(* IEC 61131-3 sources: daoli-st-library/DL_Process (part 26) *)

(* ---- FB_DL_ChamberPumpDownProfile.st ---- *)
//==============================================================================
// 功能块：FB_DL_ChamberPumpDownProfile ｜ 中文名称：腔体抽气曲线包络监视
// 所属子库：DL_Process ｜ 版本：v1.0.0 ｜ 兼容：CODESYS V3.5+ / TwinCAT 3 / 汇川 InoProShop
// 功能描述：真空腔体抽气过程包络监视——启动时锁定基线压力，以指数衰减
//           包络为参照：包络上界 p_env(t) = fBasePa x EXP(-t/tau 包络)，
//           实测压力高于上界（衰减慢于包络）持续 tSlopeTimeout → 抽速
//           异常早停（bPumpAbortReq 锁存）；滚动窗内压力样本统计（窗口
//           极差）用于判「压力停滞」（极差 < 停滞阈且未达目标真空，同
//           样归入抽速异常）。达目标真空 → 抽气完成放行（信息级）。
//           斜率判据与窗统计互为冗余：一条失效另一条仍可兜住（如压力
//           缓慢泄漏时斜率判据先报，压力卡死时停滞判据先报）。
// 遗留假设（R95 代理阈值三句）：① 代理值 = fCycleTimeS 组态扫描周期
//           [秒]（包络时间基量）；② 覆盖 0.001~0.1 秒任务周期范围；
//           ③ 覆盖不到的区间由调用方按实际任务周期重设该引脚负责，
//           该假设挂编译验证债。
// 开源溯源 (Origin)：道莅原创实现（参考真空系统抽气曲线与抽速异常判定工程惯例 分类与参数域）
// 单位表：压力[帕] / 目标真空[帕] / 包络时间常数[秒] / 时间[ms] /
//         停滞阈[帕] / 极差[帕] / 扫描周期[秒] / 样本计数[次]
// 错误码表：16#0005_01F2 信息级（抽气完成：达目标真空放行，不置
//           bError）/ 16#0005_01F3 信息级（包络逼近预警：实测压力进入
//           包络上界 1.2 倍预警带，不置 bError）/ 16#0005_0330 故障级
//           （组态非法：目标/包络/阈值域、时间窗 <= 0 或任一输入非
//           有限，置 bError）/ 16#0005_0331 故障级（抽速异常早停：斜率
//           判据或停滞判据确认，bPumpAbortReq 锁存，置 bError——该场景
//           不可由 0330 的组态类判据观测，属工艺过程独立域）/
//           16#0005_0332 故障级兜底（状态机落 ELSE，置 bError）
// 状态机：E_DL_PumpDownState（五态：eIdle=0 / ePumping=10 / eDone=20 /
//           eAbort=30 / eFault=99），CASE 含 ELSE 兜底，ELSE 置 0332 并
//           撤早停请求外的全部输出
// 边界行为：① 组态非法 → 故障态锁存，bReset 复位；② 启动拍锁定基线
//           （基线取当拍实测，非魔法数）；③ 压力非有限 → 归入抽速异常
//           域早停（0331 复用，R90：传感器数据不可信时早停为安全侧）；
//           ④ 早停锁存至 bReset；⑤ 未启动/故障态早停请求撤零并
//           bValid := FALSE（空闲态不挂请求，防误触发停泵）；⑥ 窗口
//           样本环形缓存 8 点，满窗前停滞判据不生效（样本不足不判）。
// 修订历史：v1.0.0 2026-11-17 首版（R24 派单 · ROADMAP P1 §708）
//==============================================================================

(*------------------------------------------------------------------------------
 * 枚举: E_DL_PumpDownState（归属本功能块，同文件发布，全库唯一定义）
 * 含义: 抽气监视相位，每个成员在 CASE 中有且仅有一个标签。
 *-----------------------------------------------------------------------------*)
TYPE E_DL_PumpDownState :
(
    eIdle    := 0,   // 空闲：等启动沿 / Idle, awaiting start edge
    ePumping := 10,  // 抽气：包络与停滞双判据监视 / Pumping, envelope and stagnation dual monitoring
    eDone    := 20,  // 完成：达目标真空放行 / Done, target vacuum reached
    eAbort   := 30,  // 早停：抽速异常锁存 / Abort, pumping anomaly latched
    eFault   := 99   // 故障：组态非法/非法状态 / Fault, config or illegal state
);
END_TYPE

FUNCTION_BLOCK FB_DL_ChamberPumpDownProfile
VAR_INPUT
    bStart       : BOOL;                    // 启动请求 [—]，上升沿生效 / Start request, rising edge
    bReset       : BOOL;                    // 故障复位 [—]，上升沿清锁存 / Fault reset, rising edge clears latches
    fPressPa     : LREAL;                   // 腔压实测 [帕]（绝对压力） / Chamber pressure [Pa], absolute
    fTargetPa    : LREAL := 10.0;           // 目标真空 [帕]，须 > 0 / Target vacuum [Pa], must be > 0
    fTauEnvS     : LREAL := 60.0;           // 包络时间常数 [秒]，须 > 0 / Envelope time constant [s]
    fStagThreshPa: LREAL := 0.5;            // 停滞阈 [帕]（窗极差低于此判停滞） / Stagnation threshold [Pa]
    fSlopeMargin : LREAL := 1.2;            // 包络预警带倍数 [倍]（须 >= 1） / Envelope warning margin [ratio]
    tSlopeTimeout: TIME  := T#30S;          // 抽速异常确认窗 [ms]，须 > 0 / Anomaly confirm window [ms]
    fCycleTimeS  : LREAL := 0.01;           // 任务扫描周期 [秒]，须 > 0（R95 代理阈值） / Task scan cycle [s], must be > 0, R95 proxy
END_VAR
VAR_OUTPUT
    bPumpAbortReq : BOOL;                   // 抽速异常早停请求 [—]（锁存保持） / Pump-abort request, latched
    bPumpDownDone : BOOL;                   // 抽气完成 [—]（完成态电平） / Pump-down done, completion level
    fEnvPressPa   : LREAL;                  // 包络上界 [帕]（诊断出口） / Envelope ceiling [Pa], diagnostics outlet
    eState        : E_DL_PumpDownState;     // 相位出口 [—] / Phase outlet
    eErr          : UDINT;                  // 错误码，0 = 无错，码位 16#0005_01F2 起信息级、16#0005_0330 起故障级（分带见错误码表） / Error code, 0 = no error, band info/fault per the code table
    bError        : BOOL;                   // 故障级标志，仅故障级错误置位 / Fault-class flag, set only on fault-level codes
    bValid        : BOOL;                   // 输出可用标志 / Outputs usable flag
END_VAR
VAR
    fbSlope  : TON;                         // 抽速异常确认计时（每拍无条件刷新）[ms] / Anomaly confirm timer, refreshed unconditionally
    _eState  : E_DL_PumpDownState := E_DL_PumpDownState.eIdle; // 当前相位 / Current phase
    _bCfgBad : BOOL;                        // 组态非法锁存 / Illegal config latch
    _bAbortL : BOOL;                        // 早停锁存 / Abort latch
    _bInfoDone: BOOL;                       // 完成信息当拍标志 / Done info flag of this scan
    _bInfoWarn: BOOL;                       // 预警信息当拍标志 / Warning info flag of this scan
    _fBasePa : LREAL;                       // 启动基线压力 [帕] / Startup baseline pressure [Pa]
    _fElapsedS: LREAL;                      // 抽气累计时间 [秒] / Elapsed pumping time [s]
    _afWin   : ARRAY[0..7] OF LREAL;        // 滚动窗样本环形缓存 [帕] / Rolling-window sample ring [Pa]
    _nWinIdx : INT;                         // 环形缓存写指针 [次] / Ring write index [count]
    _nWinFill: INT;                         // 环形缓存已填数 [次] / Ring fill count [count]
    _bSlopeBad: BOOL;                       // 斜率判据电平（确认窗条件） / Slope-criterion level
    _bStagBad : BOOL;                       // 停滞判据电平（确认窗条件） / Stagnation-criterion level
    _bIllegal : BOOL;                       // 非法状态标志 / Illegal state flag
    _bInit    : BOOL := FALSE;              // 首扫标志，初值 FALSE 取非判定 / First-scan flag, tested negated
END_VAR
VAR CONSTANT
    DL_CPD_INF    : LREAL := 1.7976931348623157E308; // LREAL 幅值上限 / LREAL magnitude ceiling
    DL_CPD_EPS    : LREAL := 1.0E-6;        // 浮点判零容差 [帕] / Float zero tolerance [Pa]
    DL_CPD_WIN    : INT    := 8;            // 滚动窗容量 [次] / Rolling-window capacity [count]
    DL_CPD_ZERO   : LREAL := 0.0;           // 零值常量，避免裸字面量 [混合] / Zero constant, avoids a bare literal
END_VAR
VAR
    nI       : INT;                         // 极差统计循环索引 [次] / Range-statistics loop index
    fWinHi   : LREAL;                       // 窗内最大值 [帕] / Window maximum [Pa]
    fWinLo   : LREAL;                       // 窗内最小值 [帕] / Window minimum [Pa]
END_VAR

(*------------------------------------------------------------------------------
 * 段 1｜每拍预置：早停请求先撤（安全侧；锁存态在段 6 重置），标志预清零
 *      Abort request cleared first, flags pre-cleared
 *-----------------------------------------------------------------------------*)
bPumpAbortReq := FALSE;                  // 早停请求先撤（锁存态在段 6 重置） / Abort request cleared first
bPumpDownDone := FALSE;                  // 完成电平先清 / Done level cleared first
fEnvPressPa   := DL_CPD_ZERO;            // 包络出口每拍重算 / Envelope outlet recomputed
eErr   := 16#0000_0000;                  // 错误码每拍重算 / Error code recomputed
bError := FALSE;                         // 故障标志每拍重算 / Fault flag recomputed
bValid := FALSE;                         // 可用标志每拍重算 / Usable flag recomputed
_bInfoDone := FALSE;                     // 完成信息预清零 / Done info pre-cleared
_bInfoWarn := FALSE;                     // 预警信息预清零 / Warn info pre-cleared
_bIllegal  := FALSE;                     // 非法状态预清零 / Illegal flag pre-cleared

(*------------------------------------------------------------------------------
 * 段 2｜首扫初始化
 *      First-scan initialisation
 *-----------------------------------------------------------------------------*)
IF NOT _bInit THEN
    _eState  := E_DL_PumpDownState.eIdle; // 相位空闲起步 / Phase starts idle
    _bCfgBad := FALSE;                   // 组态锁存清零 / Config latch cleared
    _bAbortL := FALSE;                   // 早停锁存清零 / Abort latch cleared
    _fElapsedS := DL_CPD_ZERO;           // 累计时间清零 / Elapsed time cleared
    _nWinIdx := 0;                       // 写指针归零 / Write index reset
    _nWinFill := 0;                      // 已填数归零 / Fill count reset
    _bInit   := TRUE;                    // 首扫只做一次 / The first scan runs once
END_IF

(*------------------------------------------------------------------------------
 * 段 3｜组态防御闸：非有限（R79）+ 目标/包络/阈值/时间窗域
 *      Configuration defense gates
 *-----------------------------------------------------------------------------*)
IF (fTargetPa <> fTargetPa) OR (ABS(fTargetPa) > DL_CPD_INF)
   OR (fTauEnvS <> fTauEnvS) OR (ABS(fTauEnvS) > DL_CPD_INF)
   OR (fStagThreshPa <> fStagThreshPa) OR (ABS(fStagThreshPa) > DL_CPD_INF)
   OR (fSlopeMargin <> fSlopeMargin) OR (ABS(fSlopeMargin) > DL_CPD_INF)
   OR (fCycleTimeS <> fCycleTimeS) OR (ABS(fCycleTimeS) > DL_CPD_INF) THEN
    _bCfgBad := TRUE;                    // 非有限归组态非法锁存 / Non-finite folded into the config latch
END_IF
IF (NOT _bCfgBad) AND ((fTargetPa <= DL_CPD_EPS) OR (fTauEnvS <= DL_CPD_EPS)
   OR (fStagThreshPa <= DL_CPD_EPS) OR (fSlopeMargin < 1.0)
   OR (tSlopeTimeout <= T#0MS) OR (fCycleTimeS <= DL_CPD_EPS)) THEN
    _bCfgBad := TRUE;                    // 目标/包络/阈值/时间窗域非法锁存 / Target, envelope, threshold and window domains latched
END_IF
IF bReset THEN
    _bCfgBad := FALSE;                   // 复位清组态锁存 / Reset clears the config latch
    _bAbortL := FALSE;                   // 复位清早停锁存 / Reset clears the abort latch
END_IF

(*------------------------------------------------------------------------------
 * 段 4｜确认窗无条件刷新（R40：CASE 之外每拍必调）
 *      Confirm timer refreshed unconditionally per R40
 *-----------------------------------------------------------------------------*)
fbSlope(IN := (_eState = E_DL_PumpDownState.ePumping)
             AND (_bSlopeBad OR _bStagBad), PT := tSlopeTimeout); // 抽速异常确认窗 / Anomaly confirm window

(*------------------------------------------------------------------------------
 * 段 5｜相位机与双判据链（CASE 含 ELSE 兜底；状态改写只出现在分支判据内，R39）
 *      Phase machine and the dual-criteria chain
 *-----------------------------------------------------------------------------*)
CASE _eState OF

    E_DL_PumpDownState.eIdle:              // 空闲：启动沿且组态合法进抽气
        IF bStart AND (NOT _bCfgBad) THEN
            _fBasePa := fPressPa;          // 基线锁定（启动拍实测，非魔法数） / Baseline locked at start
            _fElapsedS := DL_CPD_ZERO;     // 累计时间归零 / Elapsed time reset
            _nWinIdx := 0;                 // 写指针归零 / Write index reset
            _nWinFill := 0;                // 已填数归零（满窗前停滞判据不生效） / Fill reset, stagnation inert before the full window
            _eState := E_DL_PumpDownState.ePumping; // 进抽气 / To pumping
        ELSIF bStart AND _bCfgBad THEN
            _eState := E_DL_PumpDownState.eFault; // 组态非法进故障 / Illegal config to fault
        END_IF

    E_DL_PumpDownState.ePumping:           // 抽气：包络/停滞双判据 + 目标判定
        IF _bCfgBad THEN
            _eState := E_DL_PumpDownState.eFault; // 组态漂移转故障 / Config drift, fault
        ELSIF fPressPa <= fTargetPa THEN
            _bInfoDone := TRUE;            // 达目标真空（信息级，拍 N 进入） / Target vacuum reached, info
            _eState := E_DL_PumpDownState.eDone; // 本拍转出：进完成 / To done
        ELSE
            _fElapsedS := _fElapsedS + fCycleTimeS; // 累计时间推进 [秒] / Elapsed time advanced
            IF (fPressPa <> fPressPa) OR (ABS(fPressPa) > DL_CPD_INF) THEN
                _bSlopeBad := TRUE;        // 腔压非有限归抽速异常域（传感器数据不可信，早停安全侧，0331 复用 R90） / Non-finite pressure folded into the anomaly domain
            ELSE
                fEnvPressPa := _fBasePa * EXP(-_fElapsedS / fTauEnvS); // 包络上界 [帕]，分母已闸 / Envelope ceiling, denominator gated
                _bSlopeBad := fPressPa > (fSlopeMargin * fEnvPressPa); // 斜率判据：衰减慢于包络 / Slope criterion: slower than the envelope
            END_IF
            _afWin[_nWinIdx] := fPressPa;  // 样本入环 / Sample into the ring
            _nWinIdx := (_nWinIdx + 1) MOD DL_CPD_WIN; // 写指针环形推进（模 8，归一安全） / Ring index advance, modulo-normalised
            IF _nWinFill < DL_CPD_WIN THEN
                _nWinFill := _nWinFill + 1; // 已填数推进 / Fill count advanced
            END_IF
            IF _nWinFill >= DL_CPD_WIN THEN
                fWinHi := _afWin[0];       // 窗极差统计起步 / Range statistics start
                fWinLo := _afWin[0];       // 窗极差统计起步 / Range statistics start
                FOR nI := 1 TO (DL_CPD_WIN - 1) DO
                    IF _afWin[nI] > fWinHi THEN
                        fWinHi := _afWin[nI]; // 窗内最大值 / Window maximum
                    END_IF
                    IF _afWin[nI] < fWinLo THEN
                        fWinLo := _afWin[nI]; // 窗内最小值 / Window minimum
                    END_IF
                END_FOR
                _bStagBad := (fWinHi - fWinLo) < fStagThreshPa; // 停滞判据：窗极差低于阈 / Stagnation: range below the threshold
            ELSE
                _bStagBad := FALSE;        // 样本不足不判停滞（边界行为⑥） / Sample insufficient, no stagnation verdict
            END_IF
            IF fbSlope.Q THEN
                _bAbortL := TRUE;          // 抽速异常确认，早停锁存（拍 N 进入） / Anomaly confirmed, abort latched
                _eState := E_DL_PumpDownState.eAbort; // 本拍转出：进早停 / To abort
            END_IF
        END_IF

    E_DL_PumpDownState.eDone:              // 完成：等启动撤销回空闲（同拍重启防抖）
        IF NOT bStart THEN
            _eState := E_DL_PumpDownState.eIdle; // 回空闲 / Back to idle
        END_IF

    E_DL_PumpDownState.eAbort:             // 早停：请求锁存保持，bReset 才解除
        IF bReset AND (NOT _bCfgBad) THEN
            _bAbortL := FALSE;             // 复位清早停锁存 / Reset clears the abort latch
            _eState := E_DL_PumpDownState.eIdle; // 回空闲 / Back to idle
        END_IF

    E_DL_PumpDownState.eFault:             // 故障：复位沿且组态恢复回空闲
        IF bReset AND (NOT _bCfgBad) THEN
            _eState := E_DL_PumpDownState.eIdle; // 回空闲 / Back to idle
        END_IF

    ELSE                                   // 非法状态兜底（R21：CASE 必带 ELSE）
        _bIllegal := TRUE;                 // 标记非法状态 / Flag the illegal state
        _eState := E_DL_PumpDownState.eFault; // 回故障态 / Back to fault
END_CASE

IF (_eState = E_DL_PumpDownState.ePumping) AND (_fElapsedS > DL_CPD_EPS)
   AND (fPressPa > (fSlopeMargin * fEnvPressPa)) THEN
    _bInfoWarn := TRUE;                    // 包络逼近预警带（信息级） / Envelope approach warning, info
END_IF

(*------------------------------------------------------------------------------
 * 段 6｜码位出口与放行（故障级码 3 行内置 bError，R45/R101 配对）
 *      Code outlet and release, fault codes paired with bError
 *-----------------------------------------------------------------------------*)
IF _bIllegal THEN
    eErr   := 16#0005_0332;                // 故障级：状态机兜底 / Fault: state machine fallback
    bError := TRUE;                        // 置故障标志 / Raise the fault flag
ELSIF _bCfgBad THEN
    eErr   := 16#0005_0330;                // 故障级：组态非法 / Fault: illegal configuration
    bError := TRUE;                        // 置故障标志 / Raise the fault flag
ELSIF _bAbortL THEN
    eErr   := 16#0005_0331;                // 故障级：抽速异常早停锁存 / Fault: pumping anomaly, abort latched
    bError := TRUE;                        // 置故障标志 / Raise the fault flag
ELSIF _bInfoWarn THEN
    eErr := 16#0005_01F3;                  // 信息级：包络逼近预警 / Info: envelope approach warning
ELSIF _bInfoDone THEN
    eErr := 16#0005_01F2;                  // 信息级：抽气完成放行 / Info: pump-down done
END_IF

bPumpAbortReq := _bAbortL;               // 早停请求出口 = 锁存量（R99，空闲态不挂请求） / Abort outlet equals the latch
bPumpDownDone := (_eState = E_DL_PumpDownState.eDone); // 完成电平挂状态量 / Done level bound to the state
bValid := (NOT bError) AND (_eState <> E_DL_PumpDownState.eIdle); // 空闲/故障输出不可用 / Outputs unusable in idle or fault
eState := _eState;                       // 相位出口 / Phase outlet
END_FUNCTION_BLOCK

(* ---- FB_DL_ChamberPurgeDry.st ---- *)
(*
  FB_DL_ChamberPurgeDry  —  腔体干燥吹扫顺控 / Chamber purge and dry sequence control
  分类 Category : DL_Process
  码位 Code     : 16#06_0_82
  版本 Version  : 1.0.1
  溯源 Source   : OSCAT Building 语义借鉴 · clean-room 实现，仅借分类/参数域/命名，未复制源码
  修改记录 Hist : v1.0.1 2026-11-23 R75 修复——FC_DL_DewPointCalc 调用补
                  uErrorId / fVaporPa / bInRange 三出参显式回执（R73 零回执
                  挂账点修，与 VaporPressureSat 族回执口径对齐），bInRange
                  并入有效判据，主顺控逻辑零改动
  功能 Function : 1) 露点判据收敛：吹扫 → 静置 → 复测 三态循环，直到复测露点低于目标；
                  2) 三段计时各用独立 TON，且每段 IN := (在相) AND NOT ton.Q 自复位（FB33-2 硬判据）；
                  3) 复测未收敛不无限等待，超过 nMaxRetry 次即转超时态并报码。
  边界 Boundary : ① 露点入参先过有限性与物理域闸（RH 0~100 %、温度 −40~120 °C），域外不出结论；
                  ② 吹扫/静置/复测计时用三实例分段 TON，每段自复位；
                  ③ 复测超次即超时升级，不得延续吹扫无限等待；
                  ④ 超时/故障三行同向：吹扫阀关 → 干燥气阀关 → 进度标志 FALSE。
  依赖 Depends  : FC_DL_DewPointCalc（露点换算，每拍无条件调用）

  码表 Error codes（本件子码步进 16#10，避让邻件码位）:
    16#0002_0682 故障级：露点入参域外或露点函数返回无效（域闸锁存，输入恢复后自解）
    16#0002_0692 故障级：计时参数为 0 或重试上限 < 1（组态闸锁存，需 bReset 清除）
    16#0002_06A2 信息级：复测超次转超时（不置 bError，仅提示）
*)

TYPE E_DL_PurgeDryPhase :
(
    eIdle      := 0,   // 空闲 / Idle
    ePurge     := 10,  // 吹扫段 / Purge stage
    eSoak      := 20,  // 静置段 / Soak stage
    eRemeasure := 30,  // 复测段 / Re-measure stage
    eDone      := 40,  // 干燥达标 / Dry target reached
    eTimeout   := 50,  // 复测超次超时 / Retry timeout
    eFault     := 90   // 故障锁定 / Fault locked
);
END_TYPE

FUNCTION_BLOCK FB_DL_ChamberPurgeDry
VAR_INPUT
    bEnable        : BOOL;                        // 总使能，FALSE 回空闲关阀 / Master enable
    bStart         : BOOL;                        // 启动，上升沿有效 / Start, rising edge
    bReset         : BOOL;                        // 复位，上升沿清故障与超时 / Reset, clears fault and timeout
    fTempC         : REAL;                        // 腔体干球温度 [degC]，域 −40~120 / Chamber dry-bulb temperature [degC]
    fRhPct         : REAL;                        // 腔体相对湿度 [%]，域 0~100 / Chamber relative humidity [%]
    fDewTargetC    : REAL := -20.0;               // 露点目标 [degC]，复测低于此值判达标 / Dew point target [degC]
    fDewHystC      : REAL := 2.0;                 // 露点达标迟滞 [degC]，防边界抖动 / Dew point hysteresis [degC]
    tPurgeTime     : TIME := T#60S;               // 吹扫段时长 [ms]，域 > 0 / Purge stage duration
    tSoakTime      : TIME := T#30S;               // 静置段时长 [ms]，域 > 0 / Soak stage duration
    tRemeasureTime : TIME := T#20S;               // 复测段时长 [ms]，域 > 0 / Re-measure stage duration
    tDewSampleTime : TIME := T#500MS;             // 露点采样节拍 [ms]，自复位心跳 / Dew sample tick, self-resetting
    nMaxRetry      : INT := 5;                    // 最大复测次数 [次]，域 >= 1 / Max re-measure count
END_VAR
VAR_OUTPUT
    bPurgeValve    : BOOL;                        // 吹扫进气阀 [开关] / Purge inlet valve
    bDryAirValve   : BOOL;                        // 干燥气补充阀 [开关] / Dry air makeup valve
    bExhaustValve  : BOOL;                        // 排气阀 [开关] / Exhaust valve
    fDewNowC       : REAL;                        // 当前露点 [degC]，采样节拍刷新 / Current dew point [degC]
    bDewValid      : BOOL;                        // 露点有效标志 / Dew point valid flag
    nRetry         : INT;                         // 已复测次数 [次] / Re-measure count
    bInProgress    : BOOL;                        // 顺控进行中 / Sequence in progress
    bDone          : BOOL;                        // 达标完成（保持型）/ Dry done, level held
    bTimeout       : BOOL;                        // 超时标志（保持型）/ Timeout flag, level held
    bError         : BOOL;                        // 故障标志，与故障级码配对 / Fault flag paired with fault codes
    uErrorId       : UDINT;                       // 事件码，0 = 无事件 / Event code, 0 = none
    eStateOut      : E_DL_PurgeDryPhase;          // 状态机当前态，段尾单点映射 / Phase mapped at tail
END_VAR
VAR
    _eState        : E_DL_PurgeDryPhase := E_DL_PurgeDryPhase.eIdle;  // 内部状态 / Internal state
    rtrStart       : R_TRIG;                      // 启动沿 / Start edge
    rtrReset       : R_TRIG;                      // 复位沿 / Reset edge
    tonPurge       : TON;                         // 吹扫段计时（自复位）/ Purge stage timer, self-resetting
    tonSoak        : TON;                         // 静置段计时（自复位）/ Soak stage timer, self-resetting
    tonRemeasure   : TON;                         // 复测段计时（自复位）/ Re-measure stage timer
    tonDewTick     : TON;                         // 露点采样心跳（自复位）/ Dew sample tick, self-resetting
    fDewCalcC      : REAL;                        // 露点函数返回暂存 [degC] / Dew point function result
    fDewHoldC      : REAL;                        // 采样节拍锁存露点 [degC] / Latched dew point at tick
    bInputOk       : BOOL;                        // 露点入参域闸结果 / Dew input domain result
    bCfgOk         : BOOL;                        // 计时/重试组态合法 / Timer and retry configuration valid
    bConverged     : BOOL;                        // 复测收敛标志 / Convergence flag
    uFault         : UDINT;                       // 锁存故障码 / Latched fault code
    uInfo          : UDINT;                       // 信息级码 / Information code
    uDewErr        : UDINT;                       // 露点函数回执码（v1.0.1 新增接收）/ Dew point FC receipt, new in v1.0.1
    fVaporPaBuf    : REAL;                        // 露点函数水汽压回执 [Pa]（v1.0.1 新增接收，诊断）/ Dew point FC vapor pressure receipt [Pa]
    bDewInRange    : BOOL;                        // 露点函数域内回执 [-]（v1.0.1 新增接收）/ Dew point FC in-range receipt
END_VAR
VAR CONSTANT
    DL_PD_TMIN     : REAL := -40.0;               // 温度有效域下限 [degC] / Temperature domain low [degC]
    DL_PD_TMAX     : REAL := 120.0;               // 温度有效域上限 [degC] / Temperature domain high [degC]
    DL_PD_RHMIN    : REAL := 0.0;                 // 湿度有效域下限 [%] / Humidity domain low [%]
    DL_PD_RHMAX    : REAL := 100.0;               // 湿度有效域上限 [%] / Humidity domain high [%]
END_VAR

(* === 段 0 · 实例刷新（无条件周期调用，自复位节拍）=== *)
rtrStart(CLK := bStart);                          // 每拍刷新启动沿
rtrReset(CLK := bReset);                          // 每拍刷新复位沿
tonPurge(IN := (_eState = E_DL_PurgeDryPhase.ePurge) AND (NOT tonPurge.Q), PT := tPurgeTime);      // 自复位
tonSoak(IN := (_eState = E_DL_PurgeDryPhase.eSoak) AND (NOT tonSoak.Q), PT := tSoakTime);           // 自复位
tonRemeasure(IN := (_eState = E_DL_PurgeDryPhase.eRemeasure) AND (NOT tonRemeasure.Q), PT := tRemeasureTime); // 自复位
tonDewTick(IN := NOT tonDewTick.Q, PT := tDewSampleTime);                                            // 采样心跳自复位

(* === 段 1 · 域闸：入参有限性 + 物理域，域外不出结论 === *)
bInputOk := (fTempC = fTempC) AND (fRhPct = fRhPct)                          // NaN 自反判据
            AND (ABS(fTempC) < 1.0E30) AND (ABS(fRhPct) < 1.0E30)            // Inf 上限兜底
            AND (fTempC >= DL_PD_TMIN) AND (fTempC <= DL_PD_TMAX)            // 温度物理域闸
            AND (fRhPct >= DL_PD_RHMIN) AND (fRhPct <= DL_PD_RHMAX);         // 湿度物理域闸
fDewCalcC := FC_DL_DewPointCalc(fTempC := fTempC, fRhPct := fRhPct,
                                uErrorId => uDewErr, fVaporPa => fVaporPaBuf,
                                bInRange => bDewInRange);                   // 露点换算每拍无条件调用 + 三出参回执（v1.0.1）
IF bInputOk AND bDewInRange AND (fDewCalcC = fDewCalcC) AND (ABS(fDewCalcC) < 1.0E30) THEN   // 域内回执并入判据（v1.0.1）
    IF tonDewTick.Q THEN
        fDewHoldC := fDewCalcC;                   // 采样节拍到时锁存露点（每 N 时间采一次）
        bDewValid := TRUE;                        // 露点有效
    END_IF
ELSE
    bDewValid := FALSE;                           // 域外：露点无效，不清零旧值（保持诊断可读）
END_IF
bCfgOk := (tPurgeTime > T#0MS) AND (tSoakTime > T#0MS) AND (tRemeasureTime > T#0MS)
          AND (tDewSampleTime > T#0MS) AND (nMaxRetry >= 1);                 // 计时与重试组态闸
IF NOT bCfgOk THEN
    uFault := 16#0002_0692;                       // 故障级：计时参数为 0 或重试上限非法
END_IF
IF NOT bInputOk THEN
    uFault := 16#0002_0682;                       // 故障级：露点入参域外（输入恢复后段 2 自解）
END_IF
IF bInputOk AND bCfgOk THEN
    IF uFault = 16#0002_0682 THEN
        uFault := 16#0000;                        // 输入恢复即自解域闸故障（复位路径可达）
    END_IF
END_IF
IF rtrReset.Q AND bCfgOk THEN
    uFault := 16#0000;                            // 复位沿清锁存（组态已合法才允许）
END_IF

(* === 段 2 · 主状态机（ENUM + CASE，含 ELSE 兜底）=== *)
CASE _eState OF
E_DL_PurgeDryPhase.eIdle :
    nRetry := 0;                                  // 新一轮复测计数清零
    bDone := FALSE;                               // 完成标志复位
    bTimeout := FALSE;                            // 超时标志复位
    bConverged := FALSE;                          // 收敛标志复位
    uInfo := 16#0000;                             // 信息码清零（条件不满足则保持 0）
    IF uFault = 16#0002_0692 THEN
        _eState := E_DL_PurgeDryPhase.eFault;     // 组态故障优先拦截
    ELSIF rtrStart.Q THEN
        _eState := E_DL_PurgeDryPhase.ePurge;     // 本拍进入吹扫相
    END_IF

E_DL_PurgeDryPhase.ePurge :
    IF tonPurge.Q THEN
        _eState := E_DL_PurgeDryPhase.eSoak;      // 本拍行为：吹扫到时长，拍末转静置
    END_IF

E_DL_PurgeDryPhase.eSoak :
    IF tonSoak.Q THEN
        _eState := E_DL_PurgeDryPhase.eRemeasure; // 静置到时长，转复测相
    END_IF

E_DL_PurgeDryPhase.eRemeasure :
    IF tonRemeasure.Q THEN
        bConverged := bDewValid AND (fDewHoldC <= (fDewTargetC - fDewHystC));   // 露点低于目标减迟滞才判收敛
        nRetry := nRetry + 1;                     // 复测次数累加
        IF bConverged THEN
            _eState := E_DL_PurgeDryPhase.eDone;  // 收敛：转达标态
            bDone := TRUE;                        // 置位型：完成标志，段尾不清零
        ELSIF nRetry >= nMaxRetry THEN
            _eState := E_DL_PurgeDryPhase.eTimeout;   // 超次：超时升级，不无限等待
            bTimeout := TRUE;                     // 置位型：超时标志
            uInfo := 16#0002_06A2;                // 信息级：复测超次（不置 bError）
        ELSE
            _eState := E_DL_PurgeDryPhase.ePurge; // 未收敛且余次：回吹扫再循环
        END_IF
    END_IF

E_DL_PurgeDryPhase.eDone :
    bDone := TRUE;                                // 达标保持直到复位或再启动
    IF rtrStart.Q OR rtrReset.Q THEN
        _eState := E_DL_PurgeDryPhase.eIdle;      // 再启动/复位回空闲
    END_IF

E_DL_PurgeDryPhase.eTimeout :
    bTimeout := TRUE;                             // 超时标志保持，等人为处理
    IF rtrReset.Q THEN
        bTimeout := FALSE;                        // 复位沿解除超时（可到达的解除路径）
        uInfo := 16#0000;                         // 信息码同步清除
        _eState := E_DL_PurgeDryPhase.eIdle;
    END_IF

E_DL_PurgeDryPhase.eFault :
    IF (uFault = 16#0000) THEN
        _eState := E_DL_PurgeDryPhase.eIdle;      // 故障已解锁回空闲
    END_IF

ELSE
    _eState := E_DL_PurgeDryPhase.eFault;         // 非法状态拦截
    uFault := 16#0002_0692;                       // 故障级：相 ID 越界（枚举兜底路径）
END_CASE
IF NOT bEnable THEN
    _eState := E_DL_PurgeDryPhase.eIdle;          // 失能最高优先回空闲
    bInProgress := FALSE;                         // 进度标志随之为 FALSE
END_IF

(* === 段 3 · 输出映射（安全三行同向：阀门关 → 露点值 → 进度判据）=== *)
bPurgeValve   := (_eState = E_DL_PurgeDryPhase.ePurge);      // 吹扫阀仅吹扫相开
bDryAirValve  := (_eState = E_DL_PurgeDryPhase.ePurge) OR (_eState = E_DL_PurgeDryPhase.eSoak);  // 干燥气随吹扫/静置
bExhaustValve := (_eState = E_DL_PurgeDryPhase.ePurge) OR (_eState = E_DL_PurgeDryPhase.eSoak)
                 OR (_eState = E_DL_PurgeDryPhase.eRemeasure);   // 排气阀复测相亦开
IF (_eState = E_DL_PurgeDryPhase.eTimeout) OR (_eState = E_DL_PurgeDryPhase.eFault)
   OR (_eState = E_DL_PurgeDryPhase.eIdle) THEN
    bPurgeValve := FALSE;                         // 超时/故障/空闲：吹扫阀强制关
    bDryAirValve := FALSE;                        // 干燥气阀强制关
    bExhaustValve := FALSE;                       // 排气阀强制关
END_IF
fDewNowC := fDewHoldC;                            // 露点输出取采样锁存值
bInProgress := (_eState = E_DL_PurgeDryPhase.ePurge) OR (_eState = E_DL_PurgeDryPhase.eSoak)
               OR (_eState = E_DL_PurgeDryPhase.eRemeasure);   // 进度判据与阀门同向
bError := (uFault <> 16#0000);                    // 故障标志仅由故障级码置位（R45 配对）
IF bError THEN
    uErrorId := uFault;                           // 故障级优先上报
ELSE
    uErrorId := uInfo;                            // 否则上报信息级码
END_IF
eStateOut := _eState;                             // 输出枚举段尾单点映射（N2 规则）
END_FUNCTION_BLOCK

(* ---- FB_DL_ChamberTempUnitBank.st ---- *)
(*
  ==================================================================
  组件名 Component  : FB_DL_ChamberTempUnitBank
  分类   Category   : DL_Process
  版本   Version    : 1.0.0
  功能   Purpose    : 多腔室温标统一换算行。批量把 1..8 个腔室的温度实测值从
                      源温标（摄氏 / 华氏 / 开尔文）换算到目标温标，出口逐通道
                      结果、逐通道有效性掩码与统计计数。内核为「先归一到摄氏、
                      再由摄氏展开到目标温标」两段式，六种换向共用同一对归一 /
                      展开函数体，不存在重复公式分支。
  溯源   Origin     : 温标换算为公开物理定义（0 摄氏度 = 273.15 开尔文 = 32 华氏度，
                      华氏步长为摄氏的 1.8 倍）；本件为 clean-room 实现，仅借鉴来源
                      分类与参数域组织（来源标签 roadmap-p2-chamber），道莅原创设计，
                      未复制任何闭源代码行。
  平台   Platform   : 纯 IEC 61131-3（REAL / WORD / SHL 常量移位，无私有库）
  作者   Author     : 道莅代码库 · PLC 编程专家（R55）
  ------------------------------------------------------------------
  边界 Boundary     :
                      一 本件只做单位换算与有效性标记，不判工艺超温、不做滤波、不做报警；
                      二 非有限输入不穿透出口：该通道保持上拍值并置无效位；
                      三 结果低于目标温标绝对零度时按 bClampAbsZero 钳到绝对零点并置无效位；
                      四 通道游标经回钳 1..8，掩码位移量 0..7 由数组边界与循环上界共同证明；
                      五 无全局变量、无外部变量声明、无物理地址寻址。
  输出契约 Output contract:
                      afTempOut 逐通道结果；序号大于 nChamberCount 的通道保持上拍值不清零；
                      wInvalidMask 位 i-1 对应通道 i，自证向量：仅通道 1 无效 → 16#0001，
                      仅通道 8 无效 → 16#0080；
                      故障级成因 eUnitBad 与 bError 配对（R45），信息级成因永不置 bError。
  修订记录 Revision  :
    2026-11-20  v1.0.0  R55 首版（批 1 · 序号 4）
  ==================================================================
*)

TYPE E_DL_TempUnit :
(
    eCelsius    := 0,   // 摄氏度 [摄氏度] / degree Celsius
    eFahrenheit := 10,  // 华氏度 [华氏度] / degree Fahrenheit
    eKelvin     := 20   // 开尔文 [开尔文] / Kelvin
);
END_TYPE

TYPE E_DL_TubCause :
(
    eNone       := 0,   // 无成因 / no cause
    eUnitBad    := 1,   // 温标枚举非法（故障级，与 bError 配对）/ illegal temperature unit enumeration, a fault paired with bError
    eCountBad   := 2,   // 通道数越域已回钳（信息级）/ channel count out of domain and clamped, informational
    eChanBad    := 3,   // 存在非有限通道，已保持上拍值（信息级）/ non-finite channels present and held at the last value, informational
    eAbsZero    := 4    // 结果低于绝对零度已钳位（信息级）/ result below absolute zero and clamped, informational
);
END_TYPE

FUNCTION_BLOCK FB_DL_ChamberTempUnitBank
VAR_INPUT
    bEnable        : BOOL := TRUE;           // 使能，失能时全部通道保持上拍值 [-] / enable, all channels hold their last value when disabled
    bReset         : BOOL := FALSE;          // 复位上升沿清故障锁存与掩码 [-] / reset rising edge clears the fault latch and the mask
    eUnitIn        : E_DL_TempUnit := E_DL_TempUnit.eCelsius;    // 源温标 [枚举] / source temperature unit [enum]
    eUnitOut       : E_DL_TempUnit := E_DL_TempUnit.eCelsius;    // 目标温标 [枚举] / target temperature unit [enum]
    nChamberCount  : INT := 8;               // 参与换算的腔室数 [个]，域 1..8 / participating channels [count], domain 1 to 8
    bClampAbsZero  : BOOL := TRUE;           // 真 = 低于绝对零度钳位，假 = 仅置无效位不改值 [-] / true clamps below absolute zero, false only flags
END_VAR
VAR_IN_OUT
    afTempIn       : ARRAY[1..8] OF REAL;    // 逐腔室温度输入 [源温标单位]，引用型入参由调用方持有 / per chamber temperature inputs in source unit, reference parameter owned by the caller
END_VAR
VAR_OUTPUT
    afTempOut      : ARRAY[1..8] OF REAL := [8(0.0)]; // 逐腔室换算结果 [目标温标单位] / per chamber converted results in target unit
    wInvalidMask   : WORD := 16#0000;        // 无效通道掩码，位 i-1 对应通道 i [-] / invalid channel mask, bit i minus one maps to channel i
    nValidCount    : INT := 0;               // 本拍有效通道数 [个] / valid channel count of this scan
    bAllValid      : BOOL := FALSE;          // 全部参与通道有效 [-] / all participating channels valid
    bAnyInvalid    : BOOL := FALSE;          // 存在无效通道 [-] / at least one invalid channel
    fSumOut        : REAL := 0.0;            // 有效通道结果之和 [目标温标单位] / sum of the valid converted results
    fAvgOut        : REAL := 0.0;            // 有效通道结果均值 [目标温标单位] / mean of the valid converted results
    eCause         : E_DL_TubCause := E_DL_TubCause.eNone; // 成因出口 [枚举] / cause outlet [enum]
    bError         : BOOL := FALSE;          // 故障锁存标志 [-] / fault latch flag
END_VAR
VAR
    rtReset        : R_TRIG;                 // 复位沿检测，段 0 无条件刷新 / reset edge detector, refreshed unconditionally in segment zero
    _eCause        : E_DL_TubCause := E_DL_TubCause.eNone;  // 内部成因，故障级锁存、信息级每拍重算 / internal cause, latched for faults and recomputed for information
    _bFault        : BOOL := FALSE;          // 故障锁存位（温标枚举非法）/ fault latch bit for an illegal unit enumeration
    _bInit         : BOOL := FALSE;          // 首扫初始化完成标志（R310）/ first scan initialisation flag
    _bUnitInOk     : BOOL := FALSE;          // 源温标枚举合法性 [-] / source unit enumeration validity
    _bUnitOutOk    : BOOL := FALSE;          // 目标温标枚举合法性 [-] / target unit enumeration validity
    _bChanOk       : BOOL := FALSE;          // 单通道输入有限性 [-] / single channel input finiteness
    _bResultOk     : BOOL := FALSE;          // 单通道结果有限性 [-] / single channel result finiteness
    _bChanBitBad   : BOOL := FALSE;          // 单通道无效位 [-] / single channel invalid bit
    _bAbsZeroHit   : BOOL := FALSE;          // 本拍出现绝对零度钳位 [-] / an absolute zero clamp occurred this scan
    _bChanNonFin   : BOOL := FALSE;          // 本拍出现非有限通道 [-] / a non-finite channel occurred this scan
    _bCountClamped : BOOL := FALSE;          // 通道数被回钳 [-] / the channel count was clamped
    _nUseCount     : INT := 0;               // 钳定后的参与通道数 [个] / clamped participating channel count
    _nIdx          : INT := 0;               // 通道游标（1 起，回钳 1..8）[通道号] / channel cursor, one-based, clamped one through eight
    _fCelsius      : REAL := 0.0;            // 归一到摄氏度的中间量 [摄氏度] / intermediate normalised to Celsius
    _fResult       : REAL := 0.0;            // 展开到目标温标的中间量 [目标温标单位] / intermediate expanded to the target unit
    _fLowLimit     : REAL := 0.0;            // 目标温标绝对零度 [目标温标单位] / absolute zero in the target unit
    _fSum          : REAL := 0.0;            // 有效结果累加 [目标温标单位] / running sum of valid results
    _wMask         : WORD := 16#0000;        // 掩码累加器，每拍清零重建 / mask accumulator, rebuilt every scan
    _wBitOne       : WORD := 16#0001;        // 单位位常量，供常量移位使用 [-] / single bit constant for the shift
END_VAR
VAR CONSTANT
    DL_TUB_MAX        : INT := 8;            // 通道容量，同时也是游标回钳上界 [个] / channel capacity and cursor clamp upper bound
    DL_TUB_K_OFFSET   : REAL := 273.15;      // 摄氏与开尔文零点偏移 [开尔文] / zero offset between Celsius and Kelvin
    DL_TUB_F_RATIO    : REAL := 1.8;         // 华氏与摄氏步长比 [无量纲] / scale ratio between Fahrenheit and Celsius
    DL_TUB_F_OFFSET   : REAL := 32.0;        // 华氏零点偏移 [华氏度] / zero offset of Fahrenheit
    DL_TUB_ABS_C      : REAL := -273.15;     // 摄氏绝对零度 [摄氏度] / absolute zero in Celsius
    DL_TUB_ABS_F      : REAL := -459.67;     // 华氏绝对零度 [华氏度] / absolute zero in Fahrenheit
    DL_TUB_ABS_K      : REAL := 0.0;         // 开尔文绝对零度 [开尔文] / absolute zero in Kelvin
    DL_TUB_ABS_MARGIN : REAL := 0.01;        // 绝对零度容差带，吸收换算舍入 [目标温标单位] / absolute zero tolerance absorbing rounding
    DL_TUB_MASK_NONE  : WORD := 16#0000;     // 空掩码常量 [-] / empty mask constant
END_VAR

// 段 0｜复位沿无条件周期刷新（禁入分支）/ segment 0, unconditional refresh of the reset edge, never inside a branch
rtReset(CLK := bReset); // 复位沿无条件刷新 / unconditional refresh of the reset edge

// 段 1｜首扫初始化（R310）/ segment 1, first scan initialisation
IF NOT _bInit THEN // 首扫一拍 / the very first scan
    _bInit := TRUE; // 置首扫完成标志 / raise the first scan flag
    _bFault := FALSE; // 故障锁存清零 / clear the fault latch
    _eCause := E_DL_TubCause.eNone; // 成因清零 / clear the cause
    _wMask := DL_TUB_MASK_NONE; // 掩码清零 / clear the mask
    _nIdx := 1; // 游标归位 / park the cursor at one
END_IF

// 段 2｜复位沿作用域：清锁存与清成因（通道输出保持，避免读数跳变）/ segment 2, reset edge scope, the latch and cause are cleared while channel outputs are held
IF rtReset.Q THEN // 复位沿 / reset edge
    _bFault := FALSE; // 作用域一：清故障锁存 / scope one, clear the fault latch
    _eCause := E_DL_TubCause.eNone; // 作用域一：清成因 / scope one, clear the cause
    _wMask := DL_TUB_MASK_NONE; // 作用域二：清无效掩码 / scope two, clear the invalid mask
END_IF

// 段 3｜温标枚举域闸：枚举有序直比，禁枚举转整数（跨平台安全）/ segment 3, unit enumeration gate by direct comparison, never by casting an enum to an integer
_bUnitInOk := (eUnitIn = E_DL_TempUnit.eCelsius) OR (eUnitIn = E_DL_TempUnit.eFahrenheit) OR (eUnitIn = E_DL_TempUnit.eKelvin); // 源温标三选一 / the source unit is one of three
_bUnitOutOk := (eUnitOut = E_DL_TempUnit.eCelsius) OR (eUnitOut = E_DL_TempUnit.eFahrenheit) OR (eUnitOut = E_DL_TempUnit.eKelvin); // 目标温标三选一 / the target unit is one of three
IF ((NOT _bUnitInOk) OR (NOT _bUnitOutOk)) AND (NOT _bFault) THEN // 枚举非法且未锁存 / illegal enumeration and not yet latched
    _bFault := TRUE; // 置故障锁存 / raise the fault latch
    _eCause := E_DL_TubCause.eUnitBad; // 故障级成因 (R45 配对 bError) / fault grade cause paired with bError
END_IF

// 段 4｜通道数回钳：越域走信息级成因，不锁存故障 / segment 4, channel count clamping with an informational cause
_bCountClamped := FALSE; // 回钳标志预置假 / preset the clamp flag to false
_nUseCount := nChamberCount; // 通道数直通 / channel count passes through
IF _nUseCount < 1 THEN // 下越界 / below the lower bound
    _nUseCount := 1; // 回钳到 1 / clamp to one
    _bCountClamped := TRUE; // 置回钳标志 / raise the clamp flag
ELSIF _nUseCount > DL_TUB_MAX THEN // 上越界 / above the upper bound
    _nUseCount := DL_TUB_MAX; // 回钳到容量上限 / clamp to the capacity ceiling
    _bCountClamped := TRUE; // 置回钳标志 / raise the clamp flag
END_IF
IF NOT bEnable THEN // 失能：不换算，全部通道保持上拍值（R191 显式声明冻结语义）/ disabled, no conversion and every channel holds its last value
    _nUseCount := 0; // 参与通道数置零使主循环不执行 / the participating count is zeroed so the main loop does not run
END_IF

// 段 5｜目标温标绝对零度选取（三支互异，非法枚举按摄氏兜底且故障已锁存）/ segment 5, absolute zero selection for the target unit
_fLowLimit := DL_TUB_ABS_C; // 绝对零度默认取摄氏 / absolute zero defaults to Celsius
IF eUnitOut = E_DL_TempUnit.eFahrenheit THEN // 目标华氏 / target Fahrenheit
    _fLowLimit := DL_TUB_ABS_F; // 华氏绝对零度 / Fahrenheit absolute zero
ELSIF eUnitOut = E_DL_TempUnit.eKelvin THEN // 目标开尔文 / target Kelvin
    _fLowLimit := DL_TUB_ABS_K; // 开尔文绝对零度 / Kelvin absolute zero
END_IF

// 段 6｜逐通道换算主循环 / segment 6, per channel conversion loop
_wMask := DL_TUB_MASK_NONE; // 掩码每拍清零重建 / the mask is rebuilt every scan
_fSum := 0.0; // 有效结果和清零 / clear the valid result sum
nValidCount := 0; // 有效通道计数清零 / clear the valid channel count
_bAbsZeroHit := FALSE; // 绝对零度钳位标志清零 / clear the absolute zero clamp flag
_bChanNonFin := FALSE; // 非有限通道标志清零 / clear the non-finite channel flag
_nIdx := 1; // 游标自 1 起，上界由 _nUseCount 约束 / the cursor starts at one, bounded by the usable count
WHILE _nIdx <= _nUseCount DO // 循环上界为钳定后的通道数，天然不越 8 / the loop bound is the clamped count, never beyond eight
    _bChanOk := (afTempIn[_nIdx] = afTempIn[_nIdx]) AND ((afTempIn[_nIdx] - afTempIn[_nIdx]) = (afTempIn[_nIdx] - afTempIn[_nIdx])); // 输入有限性闸，NaN 用自反、无穷用差值自减 / input finiteness gate
    _bChanBitBad := FALSE; // 单通道无效位预置假 / preset the single channel invalid bit to false
    IF NOT _bChanOk THEN // 输入非有限 / non-finite input
        _bChanBitBad := TRUE; // 置该通道无效位 / raise the invalid bit of that channel
        _bChanNonFin := TRUE; // 记非有限通道成因 / record the non-finite channel cause
    ELSE
        // 段 6.1｜先归一到摄氏度 / segment 6.1, normalise to Celsius first
        IF eUnitIn = E_DL_TempUnit.eFahrenheit THEN // 源华氏 / source Fahrenheit
            _fCelsius := (afTempIn[_nIdx] - DL_TUB_F_OFFSET) / DL_TUB_F_RATIO; // 除以常量 1.8，除子为非零常量 / divided by the constant one point eight
        ELSIF eUnitIn = E_DL_TempUnit.eKelvin THEN // 源开尔文 / source Kelvin
            _fCelsius := afTempIn[_nIdx] - DL_TUB_K_OFFSET; // 减零点偏移 / subtract the zero offset
        ELSE // 源摄氏或非法枚举（故障已锁存）/ source Celsius or an illegal enumeration with the fault latched
            _fCelsius := afTempIn[_nIdx]; // 直通 / pass through
        END_IF
        // 段 6.2｜再由摄氏度展开到目标温标 / segment 6.2, expand from Celsius to the target unit
        IF eUnitOut = E_DL_TempUnit.eFahrenheit THEN // 目标华氏 / target Fahrenheit
            _fResult := _fCelsius * DL_TUB_F_RATIO + DL_TUB_F_OFFSET; // 乘步长比加零点偏移 / scale then offset
        ELSIF eUnitOut = E_DL_TempUnit.eKelvin THEN // 目标开尔文 / target Kelvin
            _fResult := _fCelsius + DL_TUB_K_OFFSET; // 加零点偏移 / add the zero offset
        ELSE // 目标摄氏或非法枚举（故障已锁存）/ target Celsius or an illegal enumeration with the fault latched
            _fResult := _fCelsius; // 直通 / pass through
        END_IF
        _bResultOk := (_fResult = _fResult) AND ((_fResult - _fResult) = (_fResult - _fResult)); // 结果有限性闸 / result finiteness gate
        IF NOT _bResultOk THEN // 结果非有限 / non-finite result
            _bChanBitBad := TRUE; // 置该通道无效位 / raise the invalid bit of that channel
            _bChanNonFin := TRUE; // 记非有限通道成因 / record the non-finite channel cause
        ELSE
            IF _fResult < (_fLowLimit + DL_TUB_ABS_MARGIN) THEN // 低于绝对零度（含舍入容差带）/ below absolute zero including the rounding band
                _bAbsZeroHit := TRUE; // 记绝对零度成因 / record the absolute zero cause
                _bChanBitBad := TRUE; // 置该通道无效位 / raise the invalid bit of that channel
                IF bClampAbsZero THEN // 需要钳位 / clamping requested
                    _fResult := _fLowLimit; // 钳到绝对零点 / clamp to absolute zero
                END_IF
            END_IF
            afTempOut[_nIdx] := _fResult; // 结果落定到该通道 / settle the result into that channel
        END_IF
        IF NOT _bChanBitBad THEN // 该通道有效 / the channel is valid
            nValidCount := nValidCount + 1; // 有效计数递增 / increment the valid count
            _fSum := _fSum + afTempOut[_nIdx]; // 累加有效结果 / accumulate the valid result
        END_IF
    END_IF
    IF _bChanBitBad THEN // 该通道无效 / the channel is invalid
        _wMask := _wMask OR SHL(_wBitOne, _nIdx - 1); // 置无效位，位移量 0..7 由数组边界与循环上界共同证明 / set the invalid bit, the shift zero through seven is proven by the array bound and the loop bound
    END_IF
    _nIdx := _nIdx + 1; // 游标递增 / increment the cursor
END_WHILE

// 段 7｜统计与成因分派（R190 归因唯一，固定优先级：故障 > 回钳 > 非有限 > 绝对零度）/ segment 7, statistics and cause dispatch with a fixed priority
bAnyInvalid := _wMask <> DL_TUB_MASK_NONE; // 存在无效通道 / at least one invalid channel
bAllValid := (_wMask = DL_TUB_MASK_NONE) AND (_nUseCount >= 1); // 全部参与通道有效 / all participating channels valid
fSumOut := _fSum; // 有效和出口 / valid sum outlet
IF nValidCount > 0 THEN // 有有效通道才可算均值 / the mean needs at least one valid channel
    fAvgOut := _fSum / INT_TO_REAL(nValidCount); // 均值，除子已证大于零 / mean, divisor proven positive
ELSE
    fAvgOut := 0.0; // 无有效通道时均值为零 / zero mean when nothing is valid
END_IF
IF _bFault THEN // 故障锁存优先 / the fault latch takes priority
    _eCause := E_DL_TubCause.eUnitBad; // 故障级成因锁存回放（禁按当下输入重推断）/ the fault cause is replayed from the latch
ELSIF _bCountClamped THEN // 通道数被回钳 / the channel count was clamped
    _eCause := E_DL_TubCause.eCountBad; // 信息级成因 / informational cause
ELSIF _bChanNonFin THEN // 存在非有限通道 / non-finite channels present
    _eCause := E_DL_TubCause.eChanBad; // 信息级成因 / informational cause
ELSIF _bAbsZeroHit THEN // 存在绝对零度钳位 / an absolute zero clamp occurred
    _eCause := E_DL_TubCause.eAbsZero; // 信息级成因 / informational cause
ELSE
    _eCause := E_DL_TubCause.eNone; // 无成因 / no cause
END_IF

// 段 8｜统一出口 / segment 8, unified outlet
wInvalidMask := _wMask; // 掩码出口 / mask outlet
eCause := _eCause; // 成因出口单点映射 / single-point cause outlet mapping
bError := _bFault; // 故障标志与锁存位同源 / the fault flag shares the latch source
END_FUNCTION_BLOCK

(* ---- FB_DL_ChangeoverSequence.st ---- *)
(*
    FB_DL_ChangeoverSequence —— 换型换产五步顺控
    ------------------------------------------------------------------
    分类      : DL_Process / Sequence
    前缀      : FB_DL_
    版本      : 1.0.1
    溯源      : T2-7 PackML（只借「最小子集 + 明确终止态」的态组织纪律，不做 17 态全集）；
                T2-8 ISA-88（只借公开条款的「配方切换需前置确认」相语义，不复制条款文本）；
                五步划分、超时策略、码位 100% 自有；clean-room 重写，未复制任何
                闭源厂商源码，参考实现仅限 MIT/Apache 许可
    平台      : 纯 IEC 61131-3，CODESYS V3.5+ / TwinCAT 3 / InoProShop 通用
    作者      : 道莅代码库 · PLC编程专家（R18）
    ------------------------------------------------------------------
    功能说明  : 把换产拆成五步可确认顺控：停机确认 → 排空清洁确认 → 配方装载确认 →
                参数下发确认 → 首件确认放行；每步独立超时，任一步确认不满足即停在该步
                等人工确认，绝不自动跳过（自动跳过是换产事故的头号成因）；
                最高危点：单步超时必须是「步内计时」，进入新步时把定时器重新装载，
                绝不能让超时沿相内累计（R40 教训复核项，本件用单拍 bStepEnter 重装）；
                超时只置信息码并记录阻塞步号，不置故障——人等确认是正常生产行为；
                放行标志只在完成态置位，失能即清零（安全侧）。
    错误码    : 16#0005_01D4 单步超时后等待人工确认（阻塞步号已记录，未置故障）——信息级，不置故障
                16#0005_01D5 预留禁用（信息级，不得挪用）
                16#0005_0302 单步超时参数非法（超时保护失效）——故障级，进故障态
                16#0005_0303 前置条件不满足（目标配方号未指定 / 确认信号缺失）——故障级，进故障态
                16#0005_0304 状态机落 ELSE 兜底（非法状态，回空闲）——用途固定，不得改作他用
    码位总账  : 16#0005_01D4 用 / 16#0005_01D5 预留 ｜ 16#0005_0302 用 / 16#0005_0303 用 / 16#0005_0304 用
    状态机    : E_DL_ChangeoverState（eIdle / eStep1 / eStep2 / eStep3 / eStep4 / eStep5 / eDone / eFault），
                CASE 含 ELSE 兜底，兜底固定置 eFault、步号 99 与 0304
    采样约定  : 三个 R_TRIG 与 fbStep 在本体首部无条件调用；bStepEnter 为单拍重装标志，
                在本体前部用后即清，进入新步时由状态迁移置位，下一拍定时器从 0 重计。
    修订记录  : 2026-11-16 v1.0.0 首次入库（R18）
                2026-11-16 v1.0.1 R18 终审修复：失能闸路径只清了内部 bReady，未清对外镜像
                bReadyForProduction，输出引脚会保留上一拍的 TRUE，违反「失能即清零」安全约定；
                已在 RETURN 前补当拍清零。对外引脚与状态机零变更。
*)

(*-----------------------------------------------------------------------------
 * 枚举: E_DL_ChangeoverState（归属本功能块，与其同文件发布）
 * 含义: 五步换产状态机离散态，步号与状态值一一对应便于 HMI 直读
 *----------------------------------------------------------------------------*)
TYPE E_DL_ChangeoverState :
(
    eIdle   := 0,      // 空闲：未启动换产 / Idle, no changeover started
    eStep1  := 10,     // 步骤一：停机确认 / Step one, machine stopped confirmation
    eStep2  := 20,     // 步骤二：排空清洁确认 / Step two, line purged and cleaned confirmation
    eStep3  := 30,     // 步骤三：配方装载确认 / Step three, recipe loaded confirmation
    eStep4  := 40,     // 步骤四：参数下发确认 / Step four, parameters applied confirmation
    eStep5  := 50,     // 步骤五：首件确认放行 / Step five, first piece released confirmation
    eDone   := 60,     // 完成：放行生产，保持到复位或中止 / Done, production released until reset or abort
    eFault  := 99      // 故障：超时参数非法 / 前置条件缺失 / 非法状态 / Fault, illegal timeout, missing precondition or an illegal state
) UINT;
END_TYPE

FUNCTION_BLOCK FB_DL_ChangeoverSequence
VAR_INPUT
    bEnable         : BOOL;                    // 使能，FALSE 回空闲并清放行 / enable, FALSE returns to idle and clears the release
    bReset          : BOOL;                    // 上升沿清故障与步序 / rising edge clears the fault and the step sequence
    bStart          : BOOL;                    // 上升沿启动换产，非空闲时忽略 / rising edge starts the changeover, ignored when not idle
    bAbort          : BOOL;                    // 上升沿中止，回空闲且不置故障 / rising edge aborts to idle without raising a fault
    uTargetRecipe   : UINT := 0;               // 目标配方号，0 表示未指定 / target recipe number, 0 means unspecified
    bMachineStopped : BOOL := FALSE;           // 步骤一确认：设备已停 / step one confirmation, the machine is stopped
    bLinePurged     : BOOL := FALSE;           // 步骤二确认：物料已排空或已清洁 / step two confirmation, the line is purged or cleaned
    bRecipeLoaded   : BOOL := FALSE;           // 步骤三确认：配方已装载且校验通过 / step three confirmation, the recipe is loaded and verified
    bParamsApplied  : BOOL := FALSE;           // 步骤四确认：参数已下发到设备层 / step four confirmation, the parameters reached the device layer
    bFirstPieceOk   : BOOL := FALSE;           // 步骤五确认：首件检验合格 / step five confirmation, the first piece passed inspection
    tStepTimeout    : TIME := T#5MIN;          // 单步超时 [ms]，范围 10 s~1 h / per step timeout [ms], range 10 s to 1 h
END_VAR
VAR_OUTPUT
    uStep              : UINT;                 // 当前步号 0 空闲 / 1~5 步 / 99 故障 / current step, 0 idle, 1~5 steps, 99 fault
    bBusy              : BOOL;                 // 换产进行中 / changeover in progress
    bDone              : BOOL;                 // 全部完成单周期脉冲 / all steps completed, single-cycle pulse
    bReadyForProduction: BOOL;                 // 放行生产，完成后保持到复位或中止 / production released, held until reset or abort
    uBlockedStep       : UINT;                 // 因超时被阻塞的步号，0 = 无 / step blocked by a timeout, 0 = none
    tStepElapsed       : TIME;                 // 当前步已耗时 [ms] / elapsed time in the current step [ms]
    eErr               : UDINT;                // 错误码，0=正常 / error id, 0=ok
    bError             : BOOL;                 // 故障标志，eErr 为故障级时 TRUE / error flag, TRUE on fault-level eErr
END_VAR
VAR
    fbTrigStart : R_TRIG;                      // 启动沿检测实例，本体首部无条件刷新 / start edge instance, refreshed unconditionally
    fbTrigReset : R_TRIG;                      // 复位沿检测实例，本体首部无条件刷新 / reset edge instance, refreshed unconditionally
    fbTrigAbort : R_TRIG;                      // 中止沿检测实例，本体首部无条件刷新 / abort edge instance, refreshed unconditionally
    fbStep      : TON;                         // 单步超时定时器，本体首部无条件刷新 / per step timeout timer, refreshed unconditionally
    eState      : E_DL_ChangeoverState := E_DL_ChangeoverState.eIdle; // 内部状态机步序 / internal state machine step
    bStepEnter  : BOOL;                        // 进入新步单拍标志，本体前部用后即清并触发定时器重装 / new step single cycle flag, consumed at the body top and triggers a timer reload
    bInStep     : BOOL;                        // 处于步一至步五之中 / inside one of the five steps
    bReady      : BOOL;                        // 放行内部保持位 / internal release holding bit
    bStepOk     : BOOL;                        // 本步确认信号成立 / the confirmation of the current step holds
    uStepInt    : UINT;                        // 内部步号寄存，对外镜像 / internal step number, mirrored to the output
    bInit       : BOOL := FALSE;               // 首扫标志，初值 FALSE，判据 NOT bInit / first-scan flag, initial FALSE, tested with NOT
END_VAR
VAR CONSTANT
    DL_CO_STEP_MAX     : UINT := 5;            // 步数上限 [步] / step count upper bound [step]
    DL_CO_TIMEOUT_MIN  : TIME := T#10S;        // 单步超时下限 [ms] / per step timeout lower bound [ms]
    DL_CO_TIMEOUT_MAX  : TIME := T#1H;         // 单步超时上限 [ms] / per step timeout upper bound [ms]
    DL_CO_STEP_FAULT   : UINT := 99;           // 故障步号 / fault step number
    DL_CO_STEP_NONE    : UINT := 0;            // 无阻塞步 / no blocked step
    DL_CO_RECIPE_NONE  : UINT := 0;            // 未指定配方号的哨兵值 / sentinel of an unspecified recipe
END_VAR

// 段 0｜输出与错误状态预置 / segment 0, preset outputs and error status
eErr := 0;                                     // 预置无错误 / preset no error
bError := FALSE;                               // 预置无故障 / preset no fault
bDone := FALSE;                                // 完成脉冲先清 / clear the done pulse first
bBusy := FALSE;                                // 预置不忙 / preset not busy

// 段 1｜首扫初始化（初值 FALSE，判据 NOT bInit）/ segment 1, first-scan initialisation
IF NOT bInit THEN
    bReady := FALSE;                           // 首扫不放行 / never release on the first scan
    uBlockedStep := DL_CO_STEP_NONE;           // 无阻塞步 / no blocked step
    uStepInt := 0;                             // 步号从 0 起 / the step starts at zero
    eState := E_DL_ChangeoverState.eIdle;      // 首扫落空闲态 / start in the idle state
    bInit := TRUE;                             // 首扫只做一次 / first scan runs once only
END_IF

// 段 2｜边沿实例无条件周期刷新（红线：严禁放入条件分支）/ segment 2, unconditional edge refresh
fbTrigStart(CLK := bStart);
fbTrigReset(CLK := bReset);
fbTrigAbort(CLK := bAbort);

// 段 3｜单步超时定时器无条件调用，随后用后即清单拍重装标志 / segment 3, unconditional timer call then consume the reload flag
bInStep := (eState = E_DL_ChangeoverState.eStep1) OR (eState = E_DL_ChangeoverState.eStep2)
        OR (eState = E_DL_ChangeoverState.eStep3) OR (eState = E_DL_ChangeoverState.eStep4)
        OR (eState = E_DL_ChangeoverState.eStep5); // 处于步一至步五 / inside one of the five steps
fbStep(IN := bInStep AND (NOT bStepEnter), PT := tStepTimeout); // 重装拍掉 IN 使 ET 归零 / the reload cycle drops the input so ET returns to zero
bStepEnter := FALSE;                           // 用后即清，绝不跨拍残留 / consumed and cleared, never leaks to the next cycle
tStepElapsed := fbStep.ET;                     // 当前步已耗时 / elapsed time in the current step

// 段 4｜超时参数闸：超时保护失效不可接受 / segment 4, timeout parameter gate
IF (tStepTimeout < DL_CO_TIMEOUT_MIN) OR (tStepTimeout > DL_CO_TIMEOUT_MAX) THEN
    eErr := 16#0005_0302;                      // 超时参数非法故障码 / illegal timeout fault id
    bError := TRUE;                            // 置故障标志 / raise the error flag
    eState := E_DL_ChangeoverState.eFault;     // 进故障态 / enter the fault state
END_IF

// 段 5｜复位与中止沿：两者都回空闲，中止不置故障（人为操作合法）/ segment 5, reset and abort return to idle, abort raises no fault
IF fbTrigReset.Q THEN
    eState := E_DL_ChangeoverState.eIdle;      // 回空闲态 / back to idle
    bReady := FALSE;                           // 撤放行 / drop the release
    uBlockedStep := DL_CO_STEP_NONE;           // 清阻塞步 / clear the blocked step
    uStepInt := 0;                             // 步号归零 / step number to zero
    bStepEnter := TRUE;                        // 定时器重装 / reload the timer
END_IF
IF fbTrigAbort.Q THEN
    eState := E_DL_ChangeoverState.eIdle;      // 中止回空闲 / abort returns to idle
    bReady := FALSE;                           // 撤放行 / drop the release
    uBlockedStep := DL_CO_STEP_NONE;           // 清阻塞步 / clear the blocked step
    uStepInt := 0;                             // 步号归零 / step number to zero
    bStepEnter := TRUE;                        // 定时器重装 / reload the timer
END_IF

// 段 6｜使能闸：失能即回空闲并撤放行（安全侧）/ segment 6, enable gate drops the release
IF NOT bEnable THEN
    eState := E_DL_ChangeoverState.eIdle;      // 回空闲态 / back to idle
    bReady := FALSE;                           // 撤放行 / drop the release
    bBusy := FALSE;                            // 不忙 / not busy
    uStep := 0;                                // 步号归零 / step number to zero
    bReadyForProduction := FALSE;              // 放行镜像当拍清零，绝不留上一拍 TRUE / clear the release mirror in the same cycle, never leak a stale TRUE
    RETURN;                                    // 失能即出口 / disabled is the exit
END_IF

// 段 7｜启动沿：仅空闲态受理 / segment 7, start edge accepted only in idle
IF fbTrigStart.Q AND (eState = E_DL_ChangeoverState.eIdle) THEN
    eState := E_DL_ChangeoverState.eStep1;     // 进第一步 / enter the first step
    uBlockedStep := DL_CO_STEP_NONE;           // 清阻塞步 / clear the blocked step
    bStepEnter := TRUE;                        // 定时器重装 / reload the timer
END_IF

// 段 8｜状态机主体（CASE 必含 ELSE 兜底，红线）/ segment 8, state machine body
CASE eState OF
    E_DL_ChangeoverState.eIdle :
        uStepInt := 0;                         // 空闲步号 0 / idle step number zero
        bBusy := FALSE;                        // 不忙 / not busy
    E_DL_ChangeoverState.eStep1 :
        uStepInt := 1;                         // 步号一 / step number one
        bBusy := TRUE;                         // 换产进行中 / changeover in progress
        IF fbStep.Q THEN
            uBlockedStep := 1;                 // 记录阻塞步 / record the blocked step
            eErr := 16#0005_01D4;              // 等待人工确认（信息级不置故障）/ waiting for manual confirmation, info level never raises a fault
        END_IF
        bStepOk := bMachineStopped;            // 本步确认 / the step confirmation
        IF bStepOk THEN
            eState := E_DL_ChangeoverState.eStep2; // 推进到下一步 / advance to the next step
            bStepEnter := TRUE;                // 定时器重装，绝不相内累计 / reload the timer, never accumulate across steps
        END_IF
    E_DL_ChangeoverState.eStep2 :
        uStepInt := 2;                         // 步号二 / step number two
        bBusy := TRUE;                         // 换产进行中 / changeover in progress
        IF fbStep.Q THEN
            uBlockedStep := 2;                 // 记录阻塞步 / record the blocked step
            eErr := 16#0005_01D4;              // 等待人工确认（信息级不置故障）/ waiting for manual confirmation, info level never raises a fault
        END_IF
        bStepOk := bMachineStopped AND bLinePurged; // 上一步完成且本步确认同时成立 / the previous step holds and this step confirms
        IF bStepOk THEN
            eState := E_DL_ChangeoverState.eStep3; // 推进到下一步 / advance to the next step
            bStepEnter := TRUE;                // 定时器重装 / reload the timer
        END_IF
    E_DL_ChangeoverState.eStep3 :
        uStepInt := 3;                         // 步号三 / step number three
        bBusy := TRUE;                         // 换产进行中 / changeover in progress
        IF uTargetRecipe = DL_CO_RECIPE_NONE THEN
            eErr := 16#0005_0303;              // 配方号未指定故障码 / unspecified recipe fault id
            bError := TRUE;                    // 置故障标志 / raise the error flag
            eState := E_DL_ChangeoverState.eFault; // 进故障态 / enter the fault state
        ELSE
            IF fbStep.Q THEN
                uBlockedStep := 3;             // 记录阻塞步 / record the blocked step
                eErr := 16#0005_01D4;          // 等待人工确认（信息级不置故障）/ waiting for manual confirmation, info level never raises a fault
            END_IF
            bStepOk := bMachineStopped AND bLinePurged AND bRecipeLoaded; // 前两步完成且配方装载确认 / the first two steps hold and the recipe is loaded
            IF bStepOk THEN
                eState := E_DL_ChangeoverState.eStep4; // 推进到下一步 / advance to the next step
                bStepEnter := TRUE;            // 定时器重装 / reload the timer
            END_IF
        END_IF
    E_DL_ChangeoverState.eStep4 :
        uStepInt := 4;                         // 步号四 / step number four
        bBusy := TRUE;                         // 换产进行中 / changeover in progress
        IF fbStep.Q THEN
            uBlockedStep := 4;                 // 记录阻塞步 / record the blocked step
            eErr := 16#0005_01D4;              // 等待人工确认（信息级不置故障）/ waiting for manual confirmation, info level never raises a fault
        END_IF
        bStepOk := bRecipeLoaded AND bParamsApplied; // 配方已装载且参数已下发 / the recipe is loaded and the parameters are applied
        IF bStepOk THEN
            eState := E_DL_ChangeoverState.eStep5; // 推进到下一步 / advance to the next step
            bStepEnter := TRUE;                // 定时器重装 / reload the timer
        END_IF
    E_DL_ChangeoverState.eStep5 :
        uStepInt := 5;                         // 步号五 / step number five
        bBusy := TRUE;                         // 换产进行中 / changeover in progress
        IF fbStep.Q THEN
            uBlockedStep := 5;                 // 记录阻塞步 / record the blocked step
            eErr := 16#0005_01D4;              // 等待人工确认（信息级不置故障）/ waiting for manual confirmation, info level never raises a fault
        END_IF
        bStepOk := bParamsApplied AND bFirstPieceOk; // 参数已下发且首件合格 / the parameters are applied and the first piece passed
        IF bStepOk THEN
            eState := E_DL_ChangeoverState.eDone; // 全部完成 / all steps completed
            bReady := TRUE;                    // 放行生产 / release production
            bDone := TRUE;                     // 完成单拍脉冲 / the single-cycle done pulse
            bBusy := FALSE;                    // 不再忙 / no longer busy
            uBlockedStep := DL_CO_STEP_NONE;   // 清阻塞步 / clear the blocked step
        END_IF
    E_DL_ChangeoverState.eDone :
        uStepInt := 6;                         // 完成步号对外按 6 表示 / the done state reports step six
        bBusy := FALSE;                        // 不忙 / not busy
        bReady := TRUE;                        // 完成态保持放行 / the done state holds the release
    E_DL_ChangeoverState.eFault :
        uStepInt := DL_CO_STEP_FAULT;          // 故障步号 99 / fault step number ninety nine
        bBusy := FALSE;                        // 不忙 / not busy
        bReady := FALSE;                       // 故障态绝不放行 / the fault state never releases production
ELSE
    eState := E_DL_ChangeoverState.eFault;     // 非法状态一律回安全故障态 / any illegal state falls back to the safe fault state
    uStepInt := DL_CO_STEP_FAULT;              // 故障步号 / the fault step number
    eErr := 16#0005_0304;                       // 本件专用兜底码，用途固定不得改作他用 / the dedicated fallback code, its purpose is fixed
    bError := TRUE;                            // 置故障标志 / raise the error flag
    bBusy := FALSE;                            // 不忙 / not busy
    bReady := FALSE;                           // 撤放行 / drop the release
END_CASE

// 段 9｜对外镜像 / segment 9, publish the mirrors
uStep := uStepInt;                             // 步号镜像 / step number mirror
bReadyForProduction := bReady;                 // 放行镜像，失能已在上方清零 / release mirror, the enable gate already cleared it above
END_FUNCTION_BLOCK

(* ---- FB_DL_ChemDosingGrav.st ---- *)
(*
  ==================================================================
  组件名 Component  : FB_DL_ChemDosingGrav
  分类   Category   : DL_Process
  版本   Version    : 1.0.0
  功能   Purpose    : 化学液定量补给称重（密度补偿外置）。按目标体积与外部注入的
                      密度算出目标质量（目标质量 = 体积 × 密度），以净重反馈判
                      定量是否达标：净重进入目标带判完成，超出上带判超量，注料相
                      超时仍在带外判欠量。密度由外部补偿模块给出，本件只做域闸与
                      质量换算，不自行推算密度。
  溯源   Origin     : 体积乘密度的质量换算与称重定量为公开工程口径；本件为
                      clean-room 实现，仅借鉴来源分类与参数域组织（来源标签
                      roadmap-p2-chemdose），道莅原创设计，未复制任何闭源代码行。
  平台   Platform   : 纯 IEC 61131-3（TON / R_TRIG / REAL 运算，无私有库）
  作者   Author     : 道莅代码库 · PLC 编程专家（R55）
  ------------------------------------------------------------------
  边界 Boundary     :
                      一 本件只做质量换算与定量判据，不驱动泵阀、不算密度（属主边界）；
                      二 密度为外置补偿输入，越域即判故障并禁止定量（防密度错致过量）；
                      三 目标质量在启动沿一次性锁存，注料期内不随引脚漂移；
                      四 净重非有限时不更新判据，出口保持上拍值；
                      五 无全局变量、无外部变量声明、无物理地址寻址。
  输出契约 Output contract:
                      fTargetMassG 在启动沿锁存，周期内不变；
                      bDoseDone 为单拍脉冲（内部位置置位、统一出口映射后撤销）；
                      bDensityOk 为密度域闸实时值，与故障锁存同源否决定量；
                      eCause 故障级成因与 bError 配对（R45），信息级永不置 bError。
  修订记录 Revision  :
    2026-11-20  v1.0.0  R55 首版（批 4 · 序号 17）
  ==================================================================
*)

TYPE E_DL_CdgState :
(
    eIdle   := 0,       // 空闲：等启动沿 / idle, waiting for the start edge
    eDose   := 10,      // 注料：净重上升中 / dosing, the net weight is rising
    eDone   := 20,      // 完成：定量判据已锁存 / done, the dosing verdict is latched
    eFault  := 90       // 故障：密度域或组态非法锁存 / fault, density or configuration out of domain
);
END_TYPE

TYPE E_DL_CdgCause :
(
    eNone       := 0,   // 无成因 / no cause
    eCfgIllegal := 1,   // 组态非法：体积、容差或时间越域（故障级，与 bError 配对）/ illegal config, volume, tolerance or time out of domain
    eDensityBad := 2,   // 密度越域或非有限，禁止定量（故障级，与 bError 配对）/ density out of domain or non-finite, dosing inhibited, a fault paired with bError
    eOverMass   := 3,   // 超量：净重越过上带（信息级，由上层决定回抽）/ over mass beyond the upper band, informational and left to the upper layer
    eUnderMass  := 4,   // 欠量：注料超时仍在带外（信息级）/ under mass after the dosing timeout, informational
    eNetBad     := 5    // 净重非有限，判据保持上拍（信息级）/ the net weight is non-finite and the verdicts hold, informational
);
END_TYPE

FUNCTION_BLOCK FB_DL_ChemDosingGrav
VAR_INPUT
    bEnable      : BOOL := TRUE;             // 使能，失能时撤命令回空闲 [-] / enable, disabling withdraws the commands and returns to idle
    bReset       : BOOL := FALSE;           // 复位上升沿清故障锁存与判据 [-] / reset rising edge clears the fault latch and the verdicts
    bStart       : BOOL := FALSE;            // 周期启动脉冲，上升沿受理 [-] / cycle start pulse, accepted on the rising edge
    fVolTargetMl : REAL := 100.0;            // 目标补给体积 [毫升]，域 大于零 / target dosing volume [millilitre], domain above zero
    fDensityKgL  : REAL := 1.2;              // 外部注入的化学液密度 [千克每升] / externally supplied chemical density [kilogram per litre]
    fDensityMinKgL : REAL := 0.5;            // 密度可接受下限 [千克每升]，域 大于零 / acceptable density floor [kilogram per litre], domain above zero
    fDensityMaxKgL : REAL := 2.5;            // 密度可接受上限 [千克每升]，须大于下限 / acceptable density ceiling [kilogram per litre], above the floor
    fNetG        : REAL := 0.0;              // 净重实测（已去皮）[克] / measured net weight, tare removed [gram]
    fTolPct      : REAL := 1.0;              // 质量容差 [百分比]，域 大于零 / mass tolerance [percent], domain above zero
    tDoseTo      : TIME := T#90S;            // 注料相超时 [毫秒]，域 大于零 / dosing phase timeout [millisecond], domain above zero
END_VAR
VAR_OUTPUT
    fTargetMassG : REAL := 0.0;              // 锁存的目标质量 [克] / latched target mass [gram]
    fDoseErrG    : REAL := 0.0;              // 净重与目标质量偏差 [克] / deviation between the net weight and the target mass [gram]
    fDosePct     : REAL := 0.0;              // 注料完成百分比 [百分比] / dosing completion ratio [percent]
    bInTol       : BOOL := FALSE;            // 净重落在质量带内 [-] / the net weight is inside the mass band
    bDensityOk   : BOOL := FALSE;            // 密度域闸通过 [-] / the density domain gate passed
    bDoseDone    : BOOL := FALSE;            // 定量完成单拍脉冲 [-] / dosing done single-shot pulse
    bOverMass    : BOOL := FALSE;            // 超量判据 [-] / over mass verdict
    bUnderMass   : BOOL := FALSE;            // 欠量判据 [-] / under mass verdict
    eState       : E_DL_CdgState := E_DL_CdgState.eIdle; // 相位出口 [枚举] / phase outlet [enum]
    eCause       : E_DL_CdgCause := E_DL_CdgCause.eNone; // 成因出口 [枚举] / cause outlet [enum]
    bError       : BOOL := FALSE;            // 故障锁存标志 [-] / fault latch flag
END_VAR
VAR
    rtStart      : R_TRIG;                   // 启动沿检测，段 0 无条件刷新 / start edge detector, refreshed unconditionally in segment zero
    rtReset      : R_TRIG;                   // 复位沿检测，段 0 无条件刷新 / reset edge detector, refreshed unconditionally in segment zero
    tonDose      : TON;                      // 注料超时，段 0 无条件刷新 / dosing timeout, refreshed unconditionally in segment zero
    _eState      : E_DL_CdgState := E_DL_CdgState.eIdle;  // 内部相位，CASE 唯一写入目标 / internal phase, the only CASE write target
    _eCause      : E_DL_CdgCause := E_DL_CdgCause.eNone;  // 信息级成因，每拍重算 / informational cause, recomputed every scan
    _eFaultCause : E_DL_CdgCause := E_DL_CdgCause.eNone;  // 故障级成因，锁存至复位沿 / fault cause, latched until the reset edge
    _bFault      : BOOL := FALSE;            // 故障锁存位 [-] / fault latch bit
    _bInit       : BOOL := FALSE;            // 首扫初始化完成标志（R310）/ first scan initialisation flag
    _bCfgBad     : BOOL := FALSE;            // 组态非法判定 [-] / illegal configuration verdict
    _bDenOk      : BOOL := FALSE;            // 密度域闸工作值 [-] / density gate working value
    _bNetOk      : BOOL := FALSE;            // 净重有限 [-] / the net weight is finite
    _bInTol      : BOOL := FALSE;            // 带内判据内部位 / internal in-target verdict
    _bOverInt    : BOOL := FALSE;            // 超量判据内部位 / internal over mass verdict
    _bUnderInt   : BOOL := FALSE;            // 欠量判据内部位 / internal under mass verdict
    _bDoneInt    : BOOL := FALSE;            // 完成脉冲内部位，统一出口映射 / internal done bit, mapped at the unified outlet
    _fTarget     : REAL := 0.0;              // 目标质量锁存值 [克] / latched target mass [gram]
    _fErr        : REAL := 0.0;              // 偏差工作值 [克] / deviation working value [gram]
    _fPct        : REAL := 0.0;              // 完成百分比工作值 [百分比] / completion ratio working value [percent]
    _fTolG       : REAL := 0.0;              // 容差绝对值 [克] / absolute tolerance [gram]
END_VAR
VAR CONSTANT
    DL_CDG_VOL_MAX   : REAL := 1.0E5;        // 体积量级上限，防量纲错配 [毫升] / volume magnitude ceiling against a mismatch [millilitre]
    DL_CDG_TOL_MAX   : REAL := 100.0;        // 容差上限 [百分比] / tolerance ceiling [percent]
    DL_CDG_MASS_MAX  : REAL := 1.0E8;        // 质量量级上限 [克] / mass magnitude ceiling [gram]
    DL_CDG_PCT_MAX   : REAL := 1000.0;       // 完成百分比上限，防目标过小放大 [百分比] / completion ratio ceiling against a tiny target
END_VAR

// 段 0｜定时器与沿检测无条件周期刷新（禁入分支），IN 只串状态闸与故障闸 / segment 0, unconditional refresh with state and fault gates on IN only
rtStart(CLK := bStart); // 启动沿无条件刷新 / unconditional refresh of the start edge
rtReset(CLK := bReset); // 复位沿无条件刷新 / unconditional refresh of the reset edge
tonDose(IN := (_eState = E_DL_CdgState.eDose) AND (NOT _bFault), PT := tDoseTo); // 注料超时，仅在注料相计时 / dosing timeout timing only in the dosing phase

// 段 1｜首扫初始化（R310）/ segment 1, first scan initialisation
IF NOT _bInit THEN // 首扫一拍 / the very first scan
    _bInit := TRUE; // 置首扫完成标志 / raise the first scan flag
    _eState := E_DL_CdgState.eIdle; // 相位从空闲起步 / the phase starts from idle
    _eCause := E_DL_CdgCause.eNone; // 信息级成因清零 / clear the informational cause
    _eFaultCause := E_DL_CdgCause.eNone; // 故障级成因清零 / clear the fault cause
    _bFault := FALSE; // 故障锁存清零 / clear the fault latch
    _fTarget := 0.0; // 目标质量清零 / clear the target mass
    _fErr := 0.0; // 偏差清零 / clear the deviation
END_IF

// 段 2｜复位沿作用域：清锁存 / 迁相位 / 清判据 / 清目标锁存 / segment 2, reset edge scope
IF rtReset.Q THEN // 复位沿 / reset edge
    _bFault := FALSE; // 作用域一：清故障锁存 / scope one, clear the fault latch
    _eFaultCause := E_DL_CdgCause.eNone; // 作用域一：清故障级成因 / scope one, clear the fault cause
    _eState := E_DL_CdgState.eIdle; // 作用域二：迁回空闲相 / scope two, migrate back to idle
    _bDoneInt := FALSE; // 作用域二：清完成脉冲内部位 / scope two, clear the internal done bit
    _bInTol := FALSE; // 作用域三：清带内判据 / scope three, clear the in-target verdict
    _bOverInt := FALSE; // 作用域三：清超量判据 / scope three, clear the over mass verdict
    _bUnderInt := FALSE; // 作用域三：清欠量判据 / scope three, clear the under mass verdict
    _fTarget := 0.0; // 作用域四：清目标质量锁存 / scope four, clear the latched target
END_IF

// 段 3｜组态域闸（R151 全覆盖）：体积、容差、密度上下限、时间 / segment 3, configuration domain gate over every pin
_bCfgBad := FALSE; // 组态非法预置假 / preset the illegal configuration verdict to false
IF (fVolTargetMl <= 0.0) OR (fVolTargetMl <> fVolTargetMl) OR (fVolTargetMl > DL_CDG_VOL_MAX) THEN // 体积越域 / the volume is out of domain
    _bCfgBad := TRUE; // 判非法 / mark illegal
END_IF
IF (fTolPct <= 0.0) OR (fTolPct > DL_CDG_TOL_MAX) OR (fTolPct <> fTolPct) THEN // 容差越域 / the tolerance is out of domain
    _bCfgBad := TRUE; // 判非法 / mark illegal
END_IF
IF (fDensityMinKgL <= 0.0) OR (fDensityMaxKgL <= fDensityMinKgL) OR (fDensityMaxKgL <> fDensityMaxKgL) THEN // 密度上下限自相矛盾 / the density bounds contradict each other
    _bCfgBad := TRUE; // 判非法 / mark illegal
END_IF
IF tDoseTo <= T#0S THEN // 注料超时非正 / the dosing timeout is not positive
    _bCfgBad := TRUE; // 判非法 / mark illegal
END_IF
IF _bCfgBad AND (NOT _bFault) THEN // 组态非法且未锁存 / illegal configuration and not yet latched
    _bFault := TRUE; // 置故障锁存 / raise the fault latch
    _eFaultCause := E_DL_CdgCause.eCfgIllegal; // 故障级成因 (R45 配对 bError) / fault grade cause paired with bError
    _eState := E_DL_CdgState.eFault; // 迁故障相 / migrate to the fault phase
END_IF

// 段 4｜密度域闸：外置补偿量越域即禁止定量（防密度错致过量）/ segment 4, density domain gate that inhibits dosing when violated
_bDenOk := (fDensityKgL = fDensityKgL) AND ((fDensityKgL - fDensityKgL) = (fDensityKgL - fDensityKgL)) AND (fDensityKgL >= fDensityMinKgL) AND (fDensityKgL <= fDensityMaxKgL); // 密度有限性与区间闸 / density finiteness and band gate
IF (NOT _bDenOk) AND (NOT _bFault) THEN // 密度越域且未锁存 / density out of domain and not yet latched
    _bFault := TRUE; // 置故障锁存 / raise the fault latch
    _eFaultCause := E_DL_CdgCause.eDensityBad; // 故障级成因 (R45 配对 bError) / fault grade cause paired with bError
    _eState := E_DL_CdgState.eFault; // 迁故障相 / migrate to the fault phase
END_IF

// 段 5｜净重闸 / segment 5, net weight gate
_eCause := E_DL_CdgCause.eNone; // 信息级成因每拍重算 / the informational cause is recomputed every scan
_bNetOk := (fNetG = fNetG) AND ((fNetG - fNetG) = (fNetG - fNetG)) AND (ABS(fNetG) <= DL_CDG_MASS_MAX); // 净重有限性与量级闸 / net weight finiteness and magnitude gate
IF (NOT _bNetOk) AND bEnable THEN // 净重非有限且使能 / the net weight is non-finite while enabled
    _eCause := E_DL_CdgCause.eNetBad; // 信息级成因 / informational cause
END_IF

// 段 6｜相位机：ENUM + CASE，含 ELSE 非法相位兜底（R128）/ segment 6, phase machine with an ELSE fallback for illegal phases
CASE _eState OF
E_DL_CdgState.eIdle: // 空闲相：等启动沿，启动沿一次性锁存目标质量 / idle, the start edge latches the target mass once
    _bInTol := FALSE; // 撤带内判据 / withdraw the in-target verdict
    _bOverInt := FALSE; // 撤超量判据 / withdraw the over mass verdict
    _bUnderInt := FALSE; // 撤欠量判据 / withdraw the under mass verdict
    IF rtStart.Q AND bEnable AND (NOT _bFault) AND _bDenOk THEN // 启动沿且使能无故障且密度可用 / start edge while enabled, unfaulted and with a usable density
        _fTarget := fVolTargetMl * fDensityKgL; // 目标质量 = 体积 × 密度，单位恰为克 / target mass equals volume times density in grams
        IF (_fTarget <> _fTarget) OR ((_fTarget - _fTarget) <> (_fTarget - _fTarget)) OR (_fTarget > DL_CDG_MASS_MAX) THEN // 目标质量非有限或超量级 / the target is non-finite or out of magnitude
            _fTarget := 0.0; // 归零，防非有限穿透判据 / zeroed so nothing non-finite reaches the verdicts
        END_IF
        _fTolG := _fTarget * fTolPct / 100.0; // 容差绝对值，除子为常量 100.0 / absolute tolerance with the constant divisor one hundred
        _eState := E_DL_CdgState.eDose; // 迁注料相 / migrate to the dosing phase
    END_IF

E_DL_CdgState.eDose: // 注料相：带内即完成，越上带判超量，超时带外判欠量 / dosing phase with three exits
    _fErr := fNetG - _fTarget; // 偏差 / deviation
    _fPct := 0.0; // 完成百分比预置零 / preset the completion ratio to zero
    IF _fTarget > 0.0 THEN // 目标可用 / the target is usable
        _fPct := fNetG / _fTarget * 100.0; // 完成百分比，除子已证大于零 / completion ratio, divisor proven positive
        IF _fPct > DL_CDG_PCT_MAX THEN // 越上限 / above the ceiling
            _fPct := DL_CDG_PCT_MAX; // 上钳 / clamp upward
        END_IF
    END_IF
    IF _bNetOk THEN // 净重可用才判据 / the verdicts need a usable net weight
        IF ABS(_fErr) <= _fTolG THEN // 落带内 / inside the band
            _bInTol := TRUE; // 置带内判据 / raise the in-target verdict
            _bDoneInt := TRUE; // 完成脉冲内部位置位（统一出口映射，R187）/ raise the internal done bit, mapped at the unified outlet
            _eState := E_DL_CdgState.eDone; // 迁完成相 / migrate to the done phase
        ELSIF _fErr > _fTolG THEN // 越过上带 / beyond the upper band
            _bOverInt := TRUE; // 置超量判据 / raise the over mass verdict
            _bInTol := FALSE; // 撤带内判据 / withdraw the in-target verdict
            _eCause := E_DL_CdgCause.eOverMass; // 信息级成因（回抽由上层决定）/ informational cause, the reclaim action belongs to the upper layer
            _eState := E_DL_CdgState.eDone; // 迁完成相（本件判据已定型）/ migrate to the done phase because the verdict is settled
        ELSIF tonDose.Q THEN // 超时仍在带外 / timed out below the band
            _bUnderInt := TRUE; // 置欠量判据 / raise the under mass verdict
            _bInTol := FALSE; // 撤带内判据 / withdraw the in-target verdict
            _eCause := E_DL_CdgCause.eUnderMass; // 信息级成因 / informational cause
            _eState := E_DL_CdgState.eDone; // 迁完成相 / migrate to the done phase
        END_IF
    ELSIF tonDose.Q THEN // 净重不可用且超时 / the net weight is unusable and the phase timed out
        _bUnderInt := TRUE; // 置欠量判据（保守侧）/ raise the under mass verdict on the conservative side
        _eState := E_DL_CdgState.eDone; // 迁完成相 / migrate to the done phase
    END_IF

E_DL_CdgState.eDone: // 完成相：判据驻留，等复位或新启动 / done phase, the verdict holds until reset or a new start
    IF rtStart.Q AND bEnable AND _bDenOk AND (NOT _bFault) THEN // 新启动沿 / a new start edge
        _fTarget := fVolTargetMl * fDensityKgL; // 目标质量重新锁存 / relatch the target mass
        _fTolG := _fTarget * fTolPct / 100.0; // 容差重算 / recompute the tolerance
        _bInTol := FALSE; // 撤带内判据 / withdraw the in-target verdict
        _bOverInt := FALSE; // 撤超量判据 / withdraw the over mass verdict
        _bUnderInt := FALSE; // 撤欠量判据 / withdraw the under mass verdict
        _eState := E_DL_CdgState.eDose; // 直接进注料相 / go straight to the dosing phase
    END_IF

E_DL_CdgState.eFault: // 故障相：判据锁存回放，等复位沿 / fault phase, the verdicts are replayed until the reset edge
    _bInTol := FALSE; // 撤带内判据 / withdraw the in-target verdict
    _bDoneInt := FALSE; // 故障拍不出完成脉冲 / no done pulse while faulted

ELSE // 非法相位兜底（R128）/ illegal phase fallback
    _bFault := TRUE; // 置故障锁存 / raise the fault latch
    _eFaultCause := E_DL_CdgCause.eCfgIllegal; // 故障级成因记组态非法 / record the illegal configuration cause
    _eState := E_DL_CdgState.eFault; // 迁故障相 / migrate to the fault phase
END_CASE

// 段 7｜失能语义：回空闲并撤完成脉冲（R191 显式声明）/ segment 7, disabled semantics
IF NOT bEnable THEN // 失能 / disabled
    _eState := E_DL_CdgState.eIdle; // 回空闲相 / return to idle
    _bDoneInt := FALSE; // 撤完成脉冲内部位 / withdraw the internal done bit
END_IF

// 段 8｜统一出口 / segment 8, unified outlet
fTargetMassG := _fTarget; // 目标质量出口（锁存量）/ target mass outlet from the latch
fDoseErrG := _fErr; // 偏差出口 / deviation outlet
fDosePct := _fPct; // 完成百分比出口 / completion ratio outlet
bInTol := _bInTol AND (NOT _bFault); // 带内出口受故障锁存否决 / the in-target outlet is vetoed by the fault latch
bOverMass := _bOverInt; // 超量出口 / over mass outlet
bUnderMass := _bUnderInt; // 欠量出口 / under mass outlet
bDensityOk := _bDenOk AND (NOT _bFault); // 密度闸出口（挂状态量）/ density gate outlet as a state quantity
bDoseDone := _bDoneInt; // 完成脉冲映射本拍值 / map the done pulse for this scan
_bDoneInt := FALSE; // 映射后立即撤销，保证单拍宽度（R187 两段式）/ revoke right after mapping to keep a single-scan width
eState := _eState; // 相位出口单点映射 / single-point phase outlet mapping
IF _bFault THEN // 故障锁存优先 / the fault latch takes priority
    eCause := _eFaultCause; // 故障级成因锁存回放 / the fault cause is replayed from the latch
ELSE
    eCause := _eCause; // 信息级成因直映 / the informational cause is mapped directly
END_IF
bError := _bFault; // 故障标志与锁存位同源 / the fault flag shares the latch source
END_FUNCTION_BLOCK

(* ---- FB_DL_ChillerApproachTrend.st ---- *)
(*

  FB_DL_ChillerApproachTrend  —  冷机逼近度趋势诊断与性能衰减预警 / Chiller approach trend and degradation early warning

  分类 Category : DL_Process

  码位 Code     : 16#06_0_95

  版本 Version  : 1.0.0

  溯源 Source   : OSCAT Building 暖通语义借鉴 · clean-room 实现，仅借分类/参数域/命名，未复制源码

  功能 Function : 1) 逼近度 = 蒸发器出水温度 − 饱和蒸发温度 [K]，滑动窗统计（复用 FB_DL_SignalStatistics）；

                  2) 趋势 = 相邻统计周期均值差折算 K/天，周期末快照对比；

                  3) 性衰预警：趋势斜率超门限带迟滞置预警，解除可达。

  边界 Boundary : ① 逼近度计算分母（换热量代理量 = 负荷率）近零时改绝对差判据（防除零）；

                  ② 负荷率低于下限冻结趋势累计并置 bFrozen（禁低负荷数据污染趋势）；

                  ③ 趋势窗样本 < 最小值不出结论；

                  ④ 预警阈值带迟滞且解除可达；

                  ⑤ 输出三行同向：逼近度 → 趋势斜率 → 预警标志。

  依赖 Depends  : FB_DL_SignalStatistics × 2（当前窗 / 上一窗均值，每拍无条件调用）

  码表 Error codes（本件子码步进 16#30 · 本格 95 与既有 9X 子码段冲突，错位至 C5/D5 避让）:

    16#0002_06C5 故障级：组态非法（周期/门限 <= 0 / 负荷率下限域非法 / 预警迟滞 <= 0）

    16#0002_06D5 故障级：相 ID 越界（枚举兜底路径）

    16#0002_06B5 信息级：输入无效本拍冻结 / 趋势窗样本不足不出结论（不置 bError）

*)

TYPE E_DL_CatPhase :

(

    eIdle   := 0,  // 空闲 / Idle

    eWatch  := 10, // 逼近度监视与趋势累计 / Approach watching and trend accumulation

    eFault  := 90  // 组态故障锁定 / Configuration fault locked

);

END_TYPE

FUNCTION_BLOCK FB_DL_ChillerApproachTrend

VAR_INPUT

    bEnable       : BOOL;                           // 总使能，FALSE 回空闲 / Master enable

    bReset        : BOOL;                           // 复位，上升沿清组态故障 / Reset, clears fault

    fChwOutC      : REAL;                           // 蒸发器出水温度 [°C] / Chilled water leaving temp [degC]

    fSatEvapC     : REAL;                           // 饱和蒸发温度 [°C] / Saturated evaporating temp [degC]

    fLoadRatePct  : REAL;                           // 负荷率 [%]（换热量代理量）/ Load rate [%], heat-transfer proxy

    fLoadLoPct    : REAL := 30.0;                   // 负荷率冻结下限 [%]，域 > 0 / Load rate freeze floor [%]

    uPeriodMin    : UINT := 60;                     // 趋势统计周期 [min]，域 > 0 / Trend period [min]

    fWarnKPerDay  : REAL := 0.5;                    // 预警斜率门限 [K/天]，域 > 0 / Warning slope threshold [K/day]

    fHystKPerDay  : REAL := 0.1;                    // 预警迟滞 [K/天]，域 > 0 / Warning hysteresis [K/day]

    fAbsDiffMaxK  : REAL := 6.0;                    // 低负荷绝对差判据门限 [K] / Low-load absolute-difference limit [K]

    fTaskCycle    : REAL := 1.0;                    // 任务周期 [s]，域 > 0 / Task cycle [s]

    fEps          : REAL := 1.0E-6;                 // 浮点判零容差 [1] / Floating zero tolerance

END_VAR

VAR_OUTPUT

    fApproachK    : REAL;                           // 当前逼近度 [K] / Current approach [K]

    fTrendKPerDay : REAL;                           // 滑动趋势 [K/天] / Sliding trend [K/day]

    bDegradWarn   : BOOL;                           // 性衰预警标志（带迟滞）/ Degradation warning flag

    bFrozen       : BOOL;                           // 低负荷/输入无效冻结标志 / Frozen by low load or invalid input

    bTrendValid   : BOOL;                           // 趋势结论有效（窗样本充足）/ Trend conclusion valid

    bError        : BOOL;                           // 故障标志，与故障级码配对 / Fault flag

    uErrorId      : UDINT;                          // 事件码，0 = 无事件 / Event code

    eStateOut     : E_DL_CatPhase;                  // 状态机当前态，段尾单点映射 / Phase mapped at tail

END_VAR

VAR

    _eState       : E_DL_CatPhase := E_DL_CatPhase.eIdle;  // 内部状态 / Internal state

    fbStatNow     : FB_DL_SignalStatistics;         // 当前窗统计实例（无条件调用）/ Current window statistics

    fbStatOld     : FB_DL_SignalStatistics;         // 上一周期快照统计实例（无条件调用）/ Previous period statistics

    rtrReset      : R_TRIG;                         // 复位沿 / Reset edge

    bCfgOk        : BOOL;                           // 组态合法标志 / Configuration valid

    bInOk         : BOOL;                           // 双温度输入本拍有效 / Both temperatures valid

    bLoadOk       : BOOL;                           // 负荷率本拍有效 / Load rate valid

    bPeriodEdge   : BOOL;                           // 周期末沿 / Period end edge

    fAccumSec     : REAL;                           // 周期累计秒 [s]（非冻结拍累计）/ Period accumulated seconds

    fMeanNowK     : REAL;                           // 当前窗逼近度均值 [K] / Current window mean [K]

    fMeanOldK     : REAL;                           // 上一周期均值快照 [K] / Previous period mean snapshot [K]

    fPeriodDay    : REAL;                           // 周期折算天 [天] / Period in days

    bSlopeUp      : BOOL;                           // 斜率越门限（电平，迟滞状态持有）/ Slope over threshold, held

    uFault        : UDINT;                          // 锁存故障码 / Latched fault code

    uInfo         : UDINT;                          // 信息级码 / Information code

END_VAR

VAR CONSTANT

    DL_CAT_INFMAX : REAL := 1.0E30;                 // 温度有限值幅值上限 [°C] / Temperature finite bound [degC]

    DL_CAT_MINWIN : INT := 8;                       // 趋势窗最小样本数 [样本] / Minimum window samples

END_VAR

(* === 段 0 · 实例刷新 === *)

rtrReset(CLK := bReset);                          // 每拍刷新复位沿

(* === 段 1 · 组态闸 === *)

bCfgOk := (UINT_TO_REAL(uPeriodMin) > fEps)               // 周期正域

          AND (fWarnKPerDay > fEps) AND (fHystKPerDay > fEps)

          AND (fLoadLoPct > fEps) AND (fLoadLoPct < 100.0)      // 负荷率下限域

          AND (fTaskCycle > fEps)

          AND (fWarnKPerDay = fWarnKPerDay) AND (fAbsDiffMaxK = fAbsDiffMaxK);  // NaN 自反

IF NOT bCfgOk THEN

    uFault := 16#0002_06C5;                       // 故障级：组态非法

END_IF

IF rtrReset.Q AND bCfgOk THEN

    uFault := 16#0000;                            // 复位沿清锁存（解除路径可达）

    bDegradWarn := FALSE;                         // 预警同步复位

    bSlopeUp := FALSE;                            // 迟滞状态复位

    fAccumSec := 0.0;                             // 周期累计清零

END_IF

uInfo := 16#0000;                                 // 信息码每拍清零

bInOk := (fChwOutC = fChwOutC) AND (ABS(fChwOutC) < DL_CAT_INFMAX)

         AND (fSatEvapC = fSatEvapC) AND (ABS(fSatEvapC) < DL_CAT_INFMAX);  // 双温度 NaN 自反 + 幅值闸

bLoadOk := (fLoadRatePct = fLoadRatePct) AND (fLoadRatePct >= 0.0) AND (fLoadRatePct <= 100.0);  // 负荷率域闸

bFrozen := (NOT bInOk) OR (NOT bLoadOk) OR (bLoadOk AND (fLoadRatePct < fLoadLoPct));  // 低负荷/无效冻结（禁污染趋势）

(* === 段 2 · 逼近度折算 === *)

fApproachK := 0.0;                                // 逼近度缺省 0

IF bInOk THEN

    fApproachK := fChwOutC - fSatEvapC;           // 逼近度 = 出水 − 饱和蒸发 [K]

END_IF

fbStatNow(fIn := fApproachK,                      // 当前窗统计（无条件调用）

          bSample := bInOk AND (NOT bFrozen),     // 冻结拍不采（低负荷数据不进窗）

          nWindow := 32,                          // 统计窗 32 样本

          bClear := rtrReset.Q);                    // 复位沿清窗

fbStatOld(fIn := fMeanNowK,                       // 上一周期统计（输入为快照均值）

          bSample := bPeriodEdge,                 // 周期末沿采一个快照

          nWindow := 8,                           // 快照窗 8 个周期

          bClear := rtrReset.Q);

IF bPeriodEdge THEN

    fMeanOldK := fMeanNowK;                       // 周期末均值快照

END_IF

(* === 段 3 · 趋势折算 === *)

bPeriodEdge := FALSE;                            // 周期沿本拍重算

IF (NOT bFrozen) AND bEnable AND (uFault = 16#0000) THEN

    fAccumSec := fAccumSec + fTaskCycle;          // 非冻结拍累计时间（暂停语义）

    IF fAccumSec >= UINT_TO_REAL(uPeriodMin) * 60.0 THEN

        bPeriodEdge := TRUE;                      // 周期末沿

        fAccumSec := 0.0;                         // 累计清零开新周期

    END_IF

END_IF

fMeanNowK := 0.0;                                 // 均值缺省 0

bTrendValid := FALSE;                             // 结论缺省无效

fTrendKPerDay := 0.0;                             // 趋势缺省 0

IF fbStatNow.bStatValid AND (fbStatNow.nCount >= DL_CAT_MINWIN) THEN

    fMeanNowK := fbStatNow.fMean;                 // 当前窗均值（样本充足才取）

    IF fbStatOld.bValid AND (fbStatOld.nCount >= 2) THEN

        fPeriodDay := UINT_TO_REAL(uPeriodMin) / 1440.0;  // 周期折算天（分母常量无除零风险）

        fTrendKPerDay := (fMeanNowK - fMeanOldK) / fPeriodDay;   // 斜率折算 K/天

        bTrendValid := TRUE;                      // 趋势结论有效

    END_IF

ELSE

    uInfo := 16#0002_06B5;                        // 信息级：趋势窗样本不足不出结论

END_IF

(* === 段 4 · 预警判定（分母近零改绝对差判据 + 迟滞）=== *)

IF bTrendValid THEN

    IF fPeriodDay > fEps THEN

        IF ABS(fTrendKPerDay) >= fWarnKPerDay THEN

            bSlopeUp := TRUE;                     // 斜率越门限（迟滞置位）

        ELSIF ABS(fTrendKPerDay) < fWarnKPerDay - fHystKPerDay THEN

            bSlopeUp := FALSE;                    // 回差带内解除（解除路径可达）

        END_IF

        bDegradWarn := bSlopeUp;                  // 预警出口

    ELSE

        (* 分母近零防御：改绝对差判据 *)

        bDegradWarn := ABS(fMeanNowK - fMeanOldK) > fAbsDiffMaxK;   // 绝对差判据（防除零）

    END_IF

ELSE

    bDegradWarn := bDegradWarn AND bTrendValid;   // 结论无效不新增预警（保持至周期更新）

END_IF

(* === 段 5 · 主状态机（ENUM + CASE，含 ELSE 兜底）=== *)

CASE _eState OF

E_DL_CatPhase.eIdle :

    IF uFault <> 16#0000 THEN

        _eState := E_DL_CatPhase.eFault;          // 故障优先

    ELSIF bEnable AND bCfgOk THEN

        _eState := E_DL_CatPhase.eWatch;          // 进监视相

    END_IF

E_DL_CatPhase.eWatch :

    IF (uFault <> 16#0000) OR (NOT bEnable) THEN

        _eState := E_DL_CatPhase.eFault;          // 故障/失能转出

    END_IF

E_DL_CatPhase.eFault :

    IF uFault = 16#0000 THEN

        _eState := E_DL_CatPhase.eIdle;           // 解锁回空闲

    END_IF

ELSE

    _eState := E_DL_CatPhase.eFault;              // 非法状态拦截

    uFault := 16#0002_06D5;                       // 故障级：相 ID 越界

END_CASE

(* === 段 6 · 输出映射 === *)

bError := (uFault <> 16#0000);                    // 故障标志仅由故障级码置位（R45 配对）

IF bError THEN

    uErrorId := uFault;                           // 故障级优先上报

ELSE

    uErrorId := uInfo;                            // 否则上报信息级码

END_IF

eStateOut := _eState;                             // 输出枚举段尾单点映射（N2 规则）

END_FUNCTION_BLOCK
